(* IEC 61131-3 sources: daoli-st-library/DL_MathData (part 25) *)

(* ---- FC_DL_StringReplaceAtEx.st ---- *)
(*
    FC_DL_StringReplaceAtEx —— 定位定长替换防御包装（与 StringReplaceAll 全局替换职责区分）
    ------------------------------------------------------------------
    分类      : DL_MathData / String
    前缀      : FC_DL_
    版本      : 1.0.0
    溯源      : IEC 61131-3 标准语义的道莅防御性实现
                （内部委托平台内建函数，外围统一错误码/钳位/双语文档；
                  未复制任何闭源厂商源码，参考实现仅限 MIT/Apache 许可）
    平台      : 纯 IEC 61131-3，CODESYS / TwinCAT / InoProShop 通用
    作者      : 道莅代码库 · PLC编程专家（R15）
    ------------------------------------------------------------------
    功能说明  : 与既有 FC_DL_StringReplaceAll（全串搜索全局替换）职责明
                确区分：本件为定位置定长覆盖——自 nPos 位序（1 基）起用
                sRep 覆盖，不搜索、不改变总长，sRep 超出串尾部分被截断。
                nPos < 1 钳 1 置 16#0001_01BD；nPos > len 原样返回置 16#0001_01BD；覆盖长
                度 = MIN(sRep 长, len-nPos+1)，sRep 被截断时按 R37 范式显
                式置 bTruncated=TRUE 与 16#0001_028B。先整串复制再覆盖（各轮带
                255 越界 EXIT 守卫），复制后显式写空字符终止符。返回值
                TRUE 表示已执行完成。
    错误码    : 0000 正常 / 16#0001_01BD 入参越界（nPos 钳位或超串长，超长时原样返回） / 16#0001_028B 上溢下溢（sRep 超串尾被截断，bTruncated=TRUE）
    修订记录  : 2026-11-16 v1.0.0 首次入库（R15）
*)
FUNCTION FC_DL_StringReplaceAtEx : BOOL
VAR_INPUT
    sIn  : STRING(255); // 源串 [字符] / source string [chars]
    sRep : STRING(255); // 覆盖串 [字符]，超串尾部分被截断 / replacement string [chars], tail beyond the source end truncated
    nPos : INT; // 覆盖起始位序 [字符位序]，1 基 / overwrite start position [char position], 1-based
END_VAR
VAR_OUTPUT
    sResult    : STRING(255); // 结果串 [字符]，总长与源串一致 / result string [chars], same length as the source
    eErr : UDINT; // 错误码，0=正常，1=位置钳位/超长，2=覆盖串截断 / error id, 0=ok, 1=position clamped or beyond length, 2=replacement truncated
    bError     : BOOL; // 是否出错，eErr 非 0 时为 TRUE / error flag, TRUE when eErr is nonzero
    bValid     : BOOL; // 输出是否有效可用 / output valid
    bTruncated : BOOL; // 截断标志，sRep 超串尾被截断时 TRUE（R37 范式） / truncation flag, TRUE when the replacement was tail-truncated
END_VAR
VAR
    nI      : INT; // 循环索引 [字符位序]，1 基 / loop index [char position], 1-based
    nLen    : INT; // 锁存的源串有效长度 [字符] / latched effective source length [chars]
    nRepLen : INT; // 锁存的覆盖串有效长度 [字符] / latched effective replacement length [chars]
    nPosC   : INT; // 钳位后的覆盖起始位序 [字符位序] / clamped overwrite start position [char position]
    nAvail  : INT; // 自起点起可用字符数 [字符] / chars available from the start position [chars]
    nUseRep : INT; // 覆盖串实际复制数 [字符] / chars actually copied from the replacement [chars]
END_VAR
VAR CONSTANT
    DL_RA_MAX : INT := 255; // 串型上限 [字符] / string type cap [chars]
END_VAR

// 段 1｜返回值与输出预置，任何早退路径不留脏码 / segment 1, preset return value and outputs
FC_DL_StringReplaceAtEx := TRUE; // 返回值预置 TRUE（已执行口径） / preset return to TRUE
sResult                 := ''; // 结果串预置空串 / preset result to the empty string
eErr                := 16#0000_0000; // 错误码预置正常 / preset error id to ok
bError                  := FALSE; // 错误标志预置无错 / preset error flag to FALSE
bValid                  := TRUE; // 有效标志预置可用 / preset valid flag to TRUE
bTruncated              := FALSE; // 截断标志预置无截断 / preset truncation flag to FALSE

// 段 2｜两串有效长度各一次锁存（空字符截止扫描 + 255 越界守卫） / segment 2, latch both effective lengths once
nI      := 1; // 索引起始 [字符位序] / index start
nLen    := 0; // 源串长度预置 [字符] / preset source length
WHILE nI <= DL_RA_MAX DO
    IF nI > DL_RA_MAX THEN    (* 越界守卫（双重保险） EN: overrun guard *)
        EXIT;
    END_IF
    IF sIn[nI] = '$00' THEN   (* 首个空字符即串结束 EN: first null char ends the string *)
        EXIT;
    END_IF
    nLen := nI; // 记录源串最后非空位序 [字符] / record the last non-null position
    nI   := nI + 1; // 每轮自增 / per-iteration increment
END_WHILE
nI      := 1; // 索引复位 / reset index
nRepLen := 0; // 覆盖串长度预置 [字符] / preset replacement length
WHILE nI <= DL_RA_MAX DO
    IF nI > DL_RA_MAX THEN    (* 越界守卫（双重保险） EN: overrun guard *)
        EXIT;
    END_IF
    IF sRep[nI] = '$00' THEN  (* 首个空字符即串结束 EN: first null char ends the string *)
        EXIT;
    END_IF
    nRepLen := nI; // 记录覆盖串最后非空位序 [字符] / record the last non-null position
    nI      := nI + 1; // 每轮自增 / per-iteration increment
END_WHILE

// 段 3｜位置闸门：nPos < 1 钳 1 置 16#0001_01BD；nPos > len 原样返回置 16#0001_01BD / segment 3, position gate, below 1 clamped to 1, beyond length returns the original with code 1
IF nPos < 1 THEN
    nPosC := 1; // 下越界钳 1 / clamped to 1
    eErr := 16#0001_01BD; // 入参越界码 / out-of-domain code
    bError   := TRUE; // 置错误标志 / raise error flag
    bValid   := FALSE; // 钳位降级 / degraded output
ELSE
    nPosC := nPos; // 域内直通 / in-domain pass-through
END_IF
IF nPosC > nLen THEN
    FOR nI := 1 TO nLen DO
        IF nI > DL_RA_MAX THEN   (* 越界守卫（双重保险） EN: overrun guard *)
            EXIT;
        END_IF
        sResult[nI] := sIn[nI]; // 位置超长原样返回 / position beyond length, original returned
    END_FOR
    IF nLen < DL_RA_MAX THEN
        sResult[nLen + 1] := '$00'; // 空字符终止符 / null terminator
    END_IF
    eErr := 16#0001_01BD; // 入参越界码（首事件优先不覆盖钳位码） / out-of-domain code, first event kept
    bError   := TRUE; // 置错误标志 / raise error flag
    bValid   := FALSE; // 输出不可用 / output invalid
    RETURN;
END_IF

// 段 4｜覆盖配额闸（R37 范式：先判定后写入，严禁静默回夹） / segment 4, overwrite quota gate, R37 paradigm, decide before writing
nAvail := nLen - nPosC + 1; // 自起点起可用字符数 [字符] / chars available from the start
IF nRepLen > nAvail THEN
    nUseRep := nAvail; // 覆盖串截到串尾 / replacement clipped to the string end
    bTruncated := TRUE; // 显式置截断标志（R37 教训） / set the truncation flag explicitly
    eErr   := 16#0001_028B; // 上溢码：sRep 超串尾已截断 / overflow code, replacement tail-truncated
    bError     := TRUE; // 置错误标志 / raise error flag
    bValid     := FALSE; // 截断降级结果 / degraded truncated output
ELSE
    nUseRep := nRepLen; // 域内直通 / in-domain pass-through
END_IF

// 段 5｜整串复制：FOR 循环 + 255 越界 EXIT 守卫 / segment 5, copy the whole source with the overrun guard
FOR nI := 1 TO nLen DO
    IF nI > DL_RA_MAX THEN       (* 越界守卫（双重保险） EN: overrun guard *)
        EXIT;
    END_IF
    sResult[nI] := sIn[nI]; // 逐字符复制 / char-by-char copy
END_FOR

// 段 6｜定长覆盖：目的位序 = nPos 起顺延，超 255 即退出 / segment 6, fixed-position overwrite
FOR nI := 1 TO nUseRep DO
    IF (nPosC + nI - 1) > DL_RA_MAX THEN   (* 目的侧越界守卫 EN: destination overrun guard *)
        EXIT;
    END_IF
    IF nI > DL_RA_MAX THEN                 (* 源侧越界守卫 EN: source overrun guard *)
        EXIT;
    END_IF
    sResult[nPosC + nI - 1] := sRep[nI]; // 逐字符覆盖 / char-by-char overwrite
END_FOR

// 段 7｜显式写终止符：总长与源串一致 / segment 7, write the terminator explicitly, total length equals the source
IF nLen < DL_RA_MAX THEN
    sResult[nLen + 1] := '$00'; // 空字符终止符 / null terminator
END_IF
END_FUNCTION

(* ---- FC_DL_StringRightEx.st ---- *)
(*
    FC_DL_StringRightEx —— 取右 n 字符防御包装（n 越界钳位 + 255 守卫逐字符复制）
    ------------------------------------------------------------------
    分类      : DL_MathData / String
    前缀      : FC_DL_
    版本      : 1.0.0
    溯源      : IEC 61131-3 标准语义的道莅防御性实现
                （内部委托平台内建函数，外围统一错误码/钳位/双语文档；
                  未复制任何闭源厂商源码，参考实现仅限 MIT/Apache 许可）
    平台      : 纯 IEC 61131-3，CODESYS / TwinCAT / InoProShop 通用
    作者      : 道莅代码库 · PLC编程专家（R15）
    ------------------------------------------------------------------
    功能说明  : 取源串右侧 nCount 个字符到 sResult。采用逐字符 FOR 复制
                （跨平台口径，不依赖平台 RIGHT 行为差异），源/目的双侧
                均带 255 越界 EXIT 守卫，复制后显式写空字符终止符。
                nCount <= 0 返回空串置 16#0001_01A6；nCount > 实际长度返回全串并
                置 16#0001_01A4（bValid=FALSE，截断诉求由错误码显式体现）。返回值
                TRUE 表示函数已执行完成，结果总在 sResult 中。
    错误码    : 0000 正常 / 16#0001_01A4 入参越界（nCount 超实际长度，已返回全串） / 16#0001_01A6 无效入参（nCount <= 0）
    修订记录  : 2026-11-16 v1.0.0 首次入库（R15）
*)
FUNCTION FC_DL_StringRightEx : BOOL
VAR_INPUT
    sIn    : STRING(255); // 源串 [字符] / source string [chars]
    nCount : INT; // 请求取右字符数 [字符]，<= 0 判无效 / requested right char count [chars], values at or below 0 invalid
END_VAR
VAR_OUTPUT
    sResult  : STRING(255); // 结果串 [字符]，右 nCount 字符 / result string [chars], right nCount chars
    eErr : UDINT; // 错误码，0=正常 / error id, 0=ok
    bError   : BOOL; // 是否出错，eErr 非 0 时为 TRUE / error flag, TRUE when eErr is nonzero
    bValid   : BOOL; // 输出是否有效可用 / output valid
END_VAR
VAR
    nI      : INT; // 循环索引 [字符位序]，1 基 / loop index [char position], 1-based
    nLen    : INT; // 锁存的源串有效长度 [字符] / latched effective source length [chars]
    nUse    : INT; // 实际复制字符数 [字符] / chars actually copied [chars]
    nSrcBgn : INT; // 源串复制起点 [字符位序] / source copy start position [char position]
END_VAR
VAR CONSTANT
    DL_RT_MAX : INT := 255; // 串型上限 [字符] / string type cap [chars]
END_VAR

// 段 1｜返回值与输出预置，任何早退路径不留脏码 / segment 1, preset return value and outputs
FC_DL_StringRightEx := TRUE; // 返回值预置 TRUE（已执行口径） / preset return to TRUE, executed semantics
sResult             := ''; // 结果串预置空串 / preset result to the empty string
eErr            := 16#0000_0000; // 错误码预置正常 / preset error id to ok
bError              := FALSE; // 错误标志预置无错 / preset error flag to FALSE
bValid              := TRUE; // 有效标志预置可用 / preset valid flag to TRUE

// 段 2｜源串有效长度一次锁存（空字符截止扫描 + 255 越界守卫） / segment 2, latch the effective source length once
nI   := 1; // 索引起始 [字符位序] / index start
nLen := 0; // 有效长度预置 [字符] / preset effective length
WHILE nI <= DL_RT_MAX DO
    IF nI > DL_RT_MAX THEN   (* 越界守卫（双重保险） EN: overrun guard, defense in depth *)
        EXIT;
    END_IF
    IF sIn[nI] = '$00' THEN  (* 首个空字符即串结束 EN: first null character marks the string end *)
        EXIT;
    END_IF
    nLen := nI; // 记录最后非空字符位序 [字符] / record the last non-null char position
    nI   := nI + 1; // 每轮自增 / per-iteration increment
END_WHILE

// 段 3｜入参域闸门：nCount <= 0 无效置 16#0001_01A6；nCount 超长度钳到全长置 16#0001_01A4 / segment 3, input domain gate
IF nCount <= 0 THEN
    sResult  := ''; // 无效入参返回空串 / invalid input returns the empty string
    eErr := 16#0001_01A6; // 无效入参码 / invalid input code
    bError   := TRUE; // 置错误标志 / raise error flag
    bValid   := FALSE; // 输出不可用 / output invalid
    RETURN;
ELSIF nCount > nLen THEN
    nUse    := nLen; // 请求超长，钳到全串长 / request beyond length, clamped to full length
    eErr := 16#0001_01A4; // 入参越界码：截断诉求显式置码 / out-of-domain code, truncation intent made explicit
    bError   := TRUE; // 置错误标志 / raise error flag
    bValid   := FALSE; // 输出为截断降级结果 / output is a degraded truncated result
ELSE
    nUse := nCount; // 域内直通 / in-domain pass-through
END_IF
nSrcBgn := nLen - nUse + 1; // 源串复制起点 = 长度减取数加一 [字符位序] / source start = length minus count plus one

// 段 4｜逐字符复制（跨平台口径）：源/目的双侧 255 越界 EXIT 守卫 / segment 4, char-by-char copy with overrun guards on both source and destination
FOR nI := 1 TO nUse DO
    IF nI > DL_RT_MAX THEN            (* 目的侧越界守卫 EN: destination overrun guard *)
        EXIT;
    END_IF
    IF (nSrcBgn + nI - 1) > DL_RT_MAX THEN   (* 源侧越界守卫 EN: source overrun guard *)
        EXIT;
    END_IF
    sResult[nI] := sIn[nSrcBgn + nI - 1]; // 逐字符复制 / char-by-char copy
END_FOR

// 段 5｜显式写终止符 / segment 5, write the terminator explicitly
IF nUse < DL_RT_MAX THEN
    sResult[nUse + 1] := '$00'; // 空字符终止符 / null terminator
END_IF
END_FUNCTION

(* ---- FC_DL_StringSplit.st ---- *)
(*==============================================================================
 * 组件名称 (Component)  : FC_DL_StringSplit
 * 所属子库 (Sublibrary) : DL_MathData
 * 当前版本 (Version)    : 1.0.0
 * 兼容性   (Platform)   : CODESYS 3.5 / TwinCAT 3 / 汇川 InoProShop / Machine Expert
 *                         仅依赖 Standard.library 的标准串函数（LEN / FIND / LEFT / DELETE）
 * 功能描述 (Function)   : 按单字符分隔符把报文拆分为字段数组。返回实际拆分出的字段数，
 *                         字段写入调用方提供的持久数组（引用型输入输出）。
 *                         采用"定位 → 取字段 → 吃掉已处理段"的标准循环，全库统一口径，
 *                         替代各项目各写一套的重复劳动（主流平台均无内置拆分函数）。
 *                         相邻分隔符产生空字段，符合 CSV 语义，不跳过、不合并；
 *                         字段数超出调用方上限时，剩余整段并入末字段并置截断标志，
 *                         结果不静默丢弃。
 * 开源溯源 (Origin)     : 原创实现。定位取段的处理范式为公开通行做法；
 *                         空字段语义与截断语义为本库差异化设计，未复制任何源码。
 * 本文件内含       : FC    FC_DL_StringSplit（单 POU，无配套类型）
 * 依赖     (Depends)    : 无 DL_ 内部依赖；Standard.library: LEN / FIND / LEFT / DELETE
 * 红线自检 (Redline)    : R1 ✓ 禁用全局存储与物理寻址 ｜ R2 ✓ 无地址直写
 *                         R3 ✓ 仅标准串函数 ｜ R4 ✓ 主循环防死锁 + 字段数钳位 + 下标双检
 *                         R5 ✓ 全变量中英双语同行注释 ｜ R6 N/A（纯函数，无状态机）
 *                         R7 N/A（无定时器/边沿实例）｜ R8 ✓ 字段上限与循环上限全常量化
 *
 * 【输出缓冲纪律 / Output buffer discipline（边界 B7，反例警告）】
 *   字段数组为引用型输入输出，调用方必须传入持久数组并在每次调用前自行清场。
 *   反例：把临时变量或每次新构造的数组传进来，上一次调用的残留字段会留在数组里，
 *   本次字段数变少时旧字段仍然可见，表现为"配方里凭空多出几个字段"的诡异故障。
 *   正确做法：一个报文一个专用数组，调用前用循环把数组元素清成空串。
 *
 * 【内存要求 / Memory requirement（边界 B10）】
 *   调用方需持有 16 × 256 字节约 4KB 的字段缓冲。单次调用最坏 16 次定位/取段/删除，
 *   无嵌套循环，耗时与报文长度呈线性关系。
 *
 * 【单字符锁定 / Single-character delimiter（边界 B1，决策 D-R2-18）】
 *   分隔符长度必须恰好为 1，否则直接拒绝且不拆分。多字符分隔会同时复杂化
 *   定位语义与截断语义，单字符已覆盖 CSV / 分号 / 竖线全部主流场景。
 *
 * 修订历史 (Revision)   :
 *   2026-11-14  v1.0.0  首版入库（Phase 1 第二轮 · Level 0 批次 A）
 *============================================================================*)
FUNCTION FC_DL_StringSplit : INT
VAR_INPUT
    sSource    : STRING(255);                 // 待拆分报文，最大 255 字符 / Source message, 255 characters max
    sDelimiter : STRING(1) := ',';            // 分隔符（单字符） / Single-character delimiter
    uMaxFields : INT := 16;                   // 最大输出字段数 [个]，合法域 1..16 / Max output fields [count], valid 1..16
END_VAR
VAR_IN_OUT
    aFields    : ARRAY[0..15] OF STRING(255); // 输出字段缓冲，调用方持有并复用 / Caller-owned reusable output buffer
END_VAR
VAR_OUTPUT
    bValid     : BOOL;                        // 拆分完整标志，FALSE = 发生截断 / Complete flag, FALSE = truncated
    uErrorId   : UDINT;                       // 故障码，0 = 无故障 / Error code, 0 = no error
END_VAR
VAR
    sTmp       : STRING(255);   // 剩余段工作副本，源串全程只读 / Working copy of the remaining segment
    nDelimPos  : INT;           // 分隔符位置（1 起始，0 = 未找到） / Delimiter position, 1-based, 0 = not found
    nFieldIdx  : INT;           // 当前字段索引 [个] / Current field index [count]
    nFieldLen  : INT;           // 当前字段长度 [字符] / Current field length [characters]
    nDelimLen  : INT;           // 分隔符长度校验值 [字符] / Delimiter length check value [characters]
    nMaxEff    : INT;           // 钳位后的最大字段数 [个] / Clamped max fields [count]
    nSrcLen    : INT;           // 源串有效长度 [字符] / Effective source length [characters]
    bRun       : BOOL;          // 循环继续标志 / Loop continuation flag
    nGuard     : DINT;          // 循环防死锁计数器 [次] / Loop deadlock guard counter [count]
    nLoop      : INT;           // 主循环索引 [次] / Main loop index [count]
END_VAR
VAR CONSTANT
    DL_SP_MAX_FIELDS : INT  := 16;   // 字段数上限 [个]，与数组维度一致 / Field cap [count], must match the array
    DL_SP_LOOP_MAX   : DINT := 64;   // 主循环防死锁上限 [次]，字段数 × 余量 / Loop guard limit [count]
    DL_SP_LEN_MAX    : INT  := 255;  // 报文字符上限 [字符]，与类型声明一致 / Message length cap [characters]
END_VAR

(*------------------------------------------------------------------------------
 * 段 1｜结果预置（P-01 范式）：先给 0 字段与成功标志
 *      Safe preset: zero fields and a success flag
 *-----------------------------------------------------------------------------*)
FC_DL_StringSplit := 0;
bValid   := TRUE;
uErrorId := 16#0000_0000;
nFieldIdx := 0;
nFieldLen := 0;
nMaxEff   := uMaxFields;

(*------------------------------------------------------------------------------
 * 段 2｜分隔符合法性（边界 B1）：长度不为 1 直接拒绝，不进入拆分流程
 *      Delimiter validity: any length other than one is rejected before splitting
 *-----------------------------------------------------------------------------*)
nDelimLen := LEN(sDelimiter);

IF nDelimLen <> 1 THEN
    bValid   := FALSE;
    uErrorId := 16#0001_0008;
    FC_DL_StringSplit := 0;
ELSE

    (*--------------------------------------------------------------------------
     * 段 3｜字段数钳位（边界 B2）：越界钳位后继续拆分，不停机
     *      Field count clamping: clamp and keep splitting, never stop the machine
     *-------------------------------------------------------------------------*)
    IF nMaxEff < 1 THEN
        nMaxEff  := 1;
        uErrorId := 16#0001_0001;
    ELSIF nMaxEff > DL_SP_MAX_FIELDS THEN
        nMaxEff  := DL_SP_MAX_FIELDS;
        uErrorId := 16#0001_0001;
    END_IF

    (* 源串长度先钳位再用：超长报文的尾部按截断处理，绝不越界读 *)
    (* Source length clamped first: an over-length message is treated as truncated *)
    nSrcLen := LEN(sSource);
    IF nSrcLen > DL_SP_LEN_MAX THEN
        nSrcLen := DL_SP_LEN_MAX;
    ELSIF nSrcLen < 0 THEN
        nSrcLen := 0;
    END_IF

    IF nSrcLen = 0 THEN
        (* 空源串是合法结果而非错误（边界 B3） *)
        (* An empty source is a legal result, not an error *)
        FC_DL_StringSplit := 0;
    ELSE

        (*----------------------------------------------------------------------
         * 段 4｜主循环（边界 B4/B5/B6）：定位、取段、删除已处理段
         *      Main loop: locate, extract, then drop the handled prefix
         *      已到最后一个可用字段而串内仍有分隔符时，剩余整段并入末字段并置截断标志
         *      On the last usable field with delimiters left, the whole remainder is kept
         *      并在置位截断标志，调用方据此识别"字段没拆完"
         *      and the truncation flag is raised so the caller can tell fields were cut
         *---------------------------------------------------------------------*)
        sTmp   := sSource;
        nLoop  := 0;
        bRun   := TRUE;
        nGuard := 0;

        WHILE bRun DO

            IF nFieldIdx >= nMaxEff THEN
                bRun := FALSE;
            ELSE
                nDelimPos := FIND(sTmp, sDelimiter);

                IF (nDelimPos > 0) AND ((nFieldIdx + 1) < nMaxEff) THEN
                    (*----------------------------------------------------------
                     * 段 4a｜常规切分：字段 = 分隔符之前的部分，然后吃掉分隔符
                     *      Normal split: the field precedes the delimiter, which is dropped
                     *      连续分隔符会自然产生长度为 0 的空字段，不跳过（边界 B6）
                     *      Consecutive delimiters yield empty fields, never skipped
                     *---------------------------------------------------------*)
                    nFieldLen := nDelimPos - 1;

                    IF nFieldLen < 0 THEN
                        nFieldLen := 0;
                    END_IF

                    IF (nFieldIdx >= 0) AND (nFieldIdx < DL_SP_MAX_FIELDS) THEN
                        aFields[nFieldIdx] := LEFT(sTmp, nFieldLen);
                    END_IF

                    sTmp      := DELETE(sTmp, nDelimPos, nDelimLen);
                    nFieldIdx := nFieldIdx + 1;

                ELSE
                    (*----------------------------------------------------------
                     * 段 4b｜末段落地：无分隔符，或已到最后一个可用字段
                     *      Final segment: no delimiter left, or the last usable field
                     *      后者若串内仍有分隔符即为截断，剩余整段并入末字段并告警
                     *      The latter with a delimiter present is a truncation and is flagged
                     *---------------------------------------------------------*)
                    IF (nFieldIdx >= 0) AND (nFieldIdx < DL_SP_MAX_FIELDS) THEN
                        aFields[nFieldIdx] := sTmp;
                    END_IF

                    nFieldIdx := nFieldIdx + 1;

                    IF nDelimPos > 0 THEN
                        bValid   := FALSE;
                        uErrorId := 16#0001_000D;
                    END_IF

                    sTmp := '';
                    bRun := FALSE;
                END_IF

            END_IF

            (* 防死锁：每轮字段索引必然递增，仍设上限兜底防止异常串函数导致死循环 *)
            (* Deadlock guard: the index always advances, the cap is a second line of defence *)
            nGuard := nGuard + 1;
            nLoop  := nLoop + 1;

            IF (nGuard > DL_SP_LOOP_MAX) OR (nLoop > DL_SP_MAX_FIELDS) THEN
                bRun     := FALSE;
                bValid   := FALSE;
                IF uErrorId = 16#0000_0000 THEN
                    uErrorId := 16#0001_0004;
                END_IF
            END_IF

        END_WHILE;

        (*----------------------------------------------------------------------
         * 段 5｜返回值：实际字段数，异常路径返回已完成的数量（P-01）
         *      Return value: the actual field count, partial counts on abnormal paths
         *---------------------------------------------------------------------*)
        IF nFieldIdx < 0 THEN
            FC_DL_StringSplit := 0;
        ELSIF nFieldIdx > DL_SP_MAX_FIELDS THEN
            FC_DL_StringSplit := DL_SP_MAX_FIELDS;
        ELSE
            FC_DL_StringSplit := nFieldIdx;
        END_IF

    END_IF
END_IF
END_FUNCTION

(* ---- FC_DL_StringStripCharsEx.st ---- *)
(*==============================================================================
 * 组件名称 (Component)  : FC_DL_StringStripCharsEx
 * 所属子库 (Sublibrary) : DL_MathData
 * 归属目录 (Directory)  : C:\Library\DL_MathData
 * 当前版本 (Version)    : 1.0.0
 * 分类/来源标签         : 函数（FUNCTION）· 纯函数 · 自定义字符集剥离
 *                         iec-std-wrapper / string / r37-reference
 * 兼容性   (Platform)   : CODESYS 3.5 / TwinCAT 3 / 汇川 InoProShop / 施耐德
 *                         Machine Expert；仅用 Standard.library 的 LEN / MID / FIND
 * 溯源声明 (Provenance) : IEC 61131-3 标准语义的道莅防御性实现——内部委托平台标准库语义，
 *                         外围统一错误码 / 钳位 / 双语注释，严禁重实现数学内核。
 * 功能一句话 (Summary)  : 去除字符串两侧属于自定义字符集的字符（区别于仅去空格的
 *                         Trim），空集输入恒等返回，全程 R37 四步长度守卫。
 *
 * 功能描述 (Function)   : LEN 一次锁存源长并与 255 比较，超限按 bAllowTrunc 分路；
 *                         合法路径用 FIND 判字符归属，从左向右收缩首界、从右向左
 *                         收缩尾界，中段一次 MID 取出，出口做长度一致性校验。
 * 与既有件边界 (Boundary): FC_DL_StringTrim 只去空格且语义固定；本件字符集是契约
 *                         参数，空串字符集即为恒等变换，不做任何猜测性补剥离。
 * 码位说明 (Codes)      : 信息 16#0002_3038 有剥离发生（nStripped 大于零）
 *                         故障 16#0002_3039 源长度域外且未允许截断（防御闸）
 *                         故障 16#0002_303A 中段取出长度与预期不一致（防御校验）
 *                         段 16#02_3_38~3B 首槽信息级、次槽起故障级。
 * 依赖说明 (Depends)    : 无 DL_ 内部依赖；仅 Standard.library 的 LEN / MID / FIND。
 * 镜像量清单 (R38)      : nSrcLen 唯一锁存量；nFirst 与 nLast 是本件的两个消费边界，
 *                         中段长度 nKeep 全部由该副本与两界导出，不重复取 LEN。
 * 红线自检 (Redline)    : 零全局依赖 ｜ 零 VAR_EXTERNAL ｜ 零 %I/%Q ｜ 纯 IEC 标准库
 *                         无除法故无除零面 ｜ 全变量双语同行注释 ｜ 无定时器实例
 * 修订历史 (Revision)   : 2026-11-18  v1.0.0  首版入库（R32 · 批 1）
 *============================================================================*)

FUNCTION FC_DL_StringStripCharsEx : BOOL
VAR_INPUT
    sSrc        : STRING(255);      // 源文本 [ASCII]，定长 255 / Source text, fixed 255 characters
    sStrip      : STRING(255);      // 剥离字符集 [ASCII]，空串即恒等 / Strip charset, empty means identity
    bAllowTrunc : BOOL := FALSE;    // 允许截断，真则截断写出，假则拒绝构造 / TRUE truncates and writes, FALSE refuses
END_VAR
VAR_OUTPUT
    sOut        : STRING(255);      // 剥离结果 [ASCII] / Stripped result
    bTruncated  : BOOL;             // 截断标志，源超上限时为真 / Set true when the source exceeded the limit
    nStripped   : INT;              // 两侧剥离的字符总数 [个] / Total characters stripped from both ends
    uErrorId    : UDINT;            // 事件码，0 表示无事件 / Event code, zero means none
END_VAR
VAR
    sMid     : STRING(255); // 中段暂存 [ASCII] / Middle segment staging
    cCh      : STRING(1);   // 当前字符 [字符] / Current character
    nSrcLen  : INT;         // 锁存的源文本长度 [字符]，R38 唯一锁存量 / Latched source length
    nFirst   : INT;         // 左边界，1 起 [索引] / Left boundary, 1-based
    nLast    : INT;         // 右边界 [索引] / Right boundary
    nKeep    : INT;         // 中段长度 [字符] / Middle segment length
    uCode    : UDINT;       // 码位暂存，出口单点写入 [码] / Code staging
END_VAR
VAR CONSTANT
    DL_STS_MAXLEN : INT := 255; // 字符串上限 [字符]，与形参声明一致 / String limit, matches the declarations
    DL_STS_ONE    : INT := 1;   // 单字符长度参数 [字符] / Single character length argument
END_VAR

(* 段 1｜输出预置与残留清除 / Pre-set and clear before any branch *)
FC_DL_StringStripCharsEx := FALSE;
sOut       := '';
sMid       := '';
bTruncated := FALSE;
nStripped  := 0;
uErrorId   := 16#0000_0000;
uCode      := 16#0000_0000;

(* 段 2｜R37 第 1 步：LEN 一次锁存 / Step one: latch the length once *)
nSrcLen := LEN(sSrc);
IF nSrcLen < 0 THEN
    nSrcLen := 0;                // 防御：异常返回值钳到零 / Defensive: clamp an anomalous result
END_IF

(* 段 3｜R37 第 2、3 步：与上限比较，超限先置标志后分路 / Compare, flag first, then branch *)
IF nSrcLen > DL_STS_MAXLEN THEN
    bTruncated := TRUE;          // 事实先记录 / Record the fact first
    IF NOT bAllowTrunc THEN
        uErrorId := 16#0002_3039; // 故障级：拒绝构造 / Fault: refuse to build
        RETURN;
    END_IF
    nSrcLen := DL_STS_MAXLEN;    // 第 4 步截断路 / Truncation path
END_IF

(* 段 4｜左界收缩：首字符属于字符集则右移 / Shrink the left boundary while the first char belongs to the set *)
nFirst := 1;
WHILE (nFirst <= nSrcLen) DO
    cCh := MID(sSrc, DL_STS_ONE, nFirst);            // 取当前首字符 / Take the current first character
    IF FIND(sStrip, cCh) > 0 THEN
        nFirst := nFirst + DL_STS_ONE;               // 属集，右移 / Belongs, shift right
    ELSE
        EXIT;                                        // 非属，停 / Not belonging, stop
    END_IF
END_WHILE

(* 段 5｜右界收缩：尾字符属于字符集则左移，越左界即停 / Shrink the right boundary, stop at the left one *)
nLast := nSrcLen;
WHILE (nLast >= nFirst) DO
    cCh := MID(sSrc, DL_STS_ONE, nLast);             // 取当前尾字符 / Take the current last character
    IF FIND(sStrip, cCh) > 0 THEN
        nLast := nLast - DL_STS_ONE;                 // 属集，左移 / Belongs, shift left
    ELSE
        EXIT;                                        // 非属，停 / Not belonging, stop
    END_IF
END_WHILE

(* 段 6｜中段一次取出：长度由两界导出，空段显式置空串 / Take the middle once; an empty segment is explicitly empty *)
nKeep := nLast - nFirst + DL_STS_ONE;                // 中段长度导出 / Derive the middle length
IF nKeep < 0 THEN
    nKeep := 0;                  // 结构性非负，仍显式兜底 / Structurally non-negative, belt and braces
END_IF
IF nKeep > 0 THEN
    sMid := MID(sSrc, nKeep, nFirst);                // 一次取出中段 / Take the middle in one shot
ELSE
    sMid := '';                  // 全串被剥离，结果空串 / Whole string stripped, result empty
END_IF

(* 段 7｜写出一致性校验（防御闸）与出口装配 / Write consistency gate and exit assembly *)
IF LEN(sMid) <> nKeep THEN
    uErrorId := 16#0002_303A;    // 故障级：取出链路异常，结果作废 / Fault: extraction chain broken
    sOut := '';
    RETURN;
END_IF
nStripped := nSrcLen - nKeep;    // 剥离计数导出 / Derive the stripped count
IF nStripped > 0 THEN
    uCode := 16#0002_3038;       // 信息级：有剥离发生 / Info: stripping happened
END_IF
sOut := sMid;
uErrorId := uCode;               // 码位单点写入 / Single write point for the code
FC_DL_StringStripCharsEx := TRUE;
END_FUNCTION

(* ---- FC_DL_StringToLowerEx.st ---- *)
(*==============================================================================
 * 组件名称 (Component)  : FC_DL_StringToLowerEx
 * 所属子库 (Sublibrary) : DL_MathData
 * 归属目录 (Directory)  : C:\Library\DL_MathData
 * 当前版本 (Version)    : 1.0.0
 * 分类/来源标签         : 函数（FUNCTION）· 纯函数 · 字符串小写扩展转换
 *                         iec-std-wrapper / string / r40-reference
 * 兼容性   (Platform)   : CODESYS 3.5 / TwinCAT 3 / 汇川 InoProShop / 施耐德
 *                         Machine Expert；仅用 Standard.library 的 LEN / MID / CONCAT / FIND
 * 溯源声明 (Provenance) : IEC 61131-3 标准语义的道莅防御性实现——内部委托平台标准库语义，
 *                         外围统一错误码 / 钳位 / 双语注释，严禁重实现数学内核。
 * 功能一句话 (Summary)  : 把 ASCII 域内大写字母映射为小写，域外字符保持原值并计数，
 *                         超长按截断标志显式分路，空串原样直通。
 * 本件存在的意义 (Why this unit exists)：
 *   各平台自带的大小写转换行为不一（有的吞掉高位字符、有的整串拒绝），本件只用
 *   标准 LEN/MID/CONCAT/FIND 做逐字符查表映射：大写字母经双码表定位转小写，
 *   其余字符原样保留并以信息码告知「有保留发生」，调用方永远知道结果里混了什么。
 * 功能描述 (Function)   : 第 1 步 LEN 一次锁存源长；第 2 步与 255 上限比较；第 3 步
 *                         超限先置截断标志（255 上限显式化，不依赖平台隐式截断）；
 *                         第 4 步按 bAllowTrunc 分路截断写出或拒绝。
 *                         空串直通：源长为 0 时不进循环、写出计数 0 等于源长 0，
 *                         出口装配返回 TRUE 且不占任何码位。
 *                         合法路径逐字符取字符：落在 'A'..'Z' 域内的用 FIND 在大写
 *                         码表定位后到同位小写码表取字符，域外字符保持并累计 nKept。
 * 与既有件边界 (Boundary): 本件为 FC_DL_StringToUpperEx 的严格对偶件（映射方向互逆、
 *                         四步样板与分路口径逐条对应），只做 ASCII A..Z 域内映射，
 *                         不做 Unicode 与本地化。
 * 码位说明 (Codes)      : 信息 16#0001_0499 源超 255 上限，已按上限截断写出
 *                         故障 16#0001_03D4 源超上限且未允许截断（防御闸拒绝）
 *                         故障 16#0001_03D5 写出计数与源长不一致（防御校验）
 *                         （R90 反证句：截断事实无法由 sDst 观测——截断与正常写出
 *                           结果均为合法串且返回值同为 TRUE，故截断侧须占码；
 *                           计数不一致属写出链路异常，与截断、保留场景的输出组合
 *                           （空串加故障码）均不同，故独立占码）
 * 依赖说明 (Depends)    : 无 DL_ 内部依赖；仅 Standard.library 的 LEN / MID / CONCAT / FIND。
 * 镜像量清单 (R38)      : nSrcLen 是本件唯一锁存量，入口一次导出，其后比较与循环
 *                         上界全部读该副本，全文不再对入参串取长度。
 * 遗留假设 (Legacy)     : 字符比较使用 >= / <= 排序比较（与库内 FC_DL_StringToUpperEx
 *                         同口径）；若某平台未实现 STRING 排序比较，须在编译门槛里
 *                         核对后改走 FIND 查表判定。
 * 红线自检 (Redline)    : 零全局依赖 ｜ 零 VAR_EXTERNAL ｜ 零 %I/%Q ｜ 纯 IEC 标准库
 *                         无除法故无除零面 ｜ 全变量双语同行注释 ｜ 无定时器实例
 * 修订历史 (Revision)   : 2026-11-19  v1.0.0  首版入库（R40 · 批 3 · T0 快车道）
 *============================================================================*)

FUNCTION FC_DL_StringToLowerEx : BOOL
VAR_INPUT
    sSrc        : STRING(255);      // 源文本 [ASCII]，定长 255 ｜ source text, fixed 255 characters
    bAllowTrunc : BOOL := FALSE;    // 允许截断，真则截断写出，假则拒绝构造 ｜ TRUE truncates and writes, FALSE refuses
END_VAR
VAR_OUTPUT
    sDst        : STRING(255);      // 小写结果 [ASCII]，域外字符保持原值 ｜ lowercase result, out-of-domain chars kept
    bTruncated  : BOOL;             // 截断标志，源超上限时为真 ｜ set true when the source exceeded the limit
    nKept       : INT;              // 保持原值的域外字符个数 [个] ｜ count of kept out-of-domain characters
    uErrorId    : UDINT;            // 事件码，0 表示无事件 ｜ event code, zero means none
END_VAR
VAR
    sTmp     : STRING(255); // 结果累积缓冲 [ASCII]，出口一次性赋给 sDst ｜ result staging buffer, assigned to sDst once at the exit
    cCh      : STRING(1);   // 当前字符 [字符] ｜ current character
    sLo      : STRING(1);   // 转换后的字符 [字符] ｜ converted character
    nPos     : INT;         // 字符在码表中的位置 [索引]，1 起 ｜ character position in the code table, 1-based
    nSrcLen  : INT;         // 锁存的源文本长度 [字符]，本件唯一锁存量 ｜ latched source length, the single latched quantity
    nWritten : INT;         // 写出计数 [字符]，出口与 nSrcLen 比对 ｜ written count compared at the exit
    uCode    : UDINT;       // 码位暂存，出口单点写入 [码] ｜ code staging, written once at the exit
END_VAR
VAR CONSTANT
    DL_STL_MAXLEN : INT := 255; // 字符串上限 [字符]，与形参声明一致 ｜ string limit, matches the declarations
    DL_STL_ONE    : INT := 1;   // 单字符长度参数 [字符] ｜ single character length argument
END_VAR

// 段 1｜输出预置与残留清除：先清空再分流，拒绝路不露旧值 ｜ preset and clear before any branch, the refusal path exposes no stale value
FC_DL_StringToLowerEx := FALSE; // 预置返回失败 ｜ preset return FALSE
sDst       := '';        // 结果清空 ｜ clear the result
sTmp       := '';        // 暂存清空 ｜ clear the staging buffer
bTruncated := FALSE;     // 截断标志清零 ｜ clear the truncation flag
nKept      := 0;         // 保留计数清零 ｜ clear the kept count
nWritten   := 0;         // 写出计数清零 ｜ clear the written count
uErrorId   := 16#0000_0000; // 事件码清零 ｜ clear the event code
uCode      := 16#0000_0000; // 码位暂存清零 ｜ clear the code staging

// 段 2｜LEN 一次锁存 ｜ latch the length once
nSrcLen := LEN(sSrc);        // 源长只取一次，循环内禁重复 LEN ｜ latch the length once, never call LEN again in the loop
IF nSrcLen < 0 THEN
    nSrcLen := 0;            // 防御：异常返回值钳到零 ｜ defensive: clamp an anomalous result to zero
END_IF

// 段 3｜与上限比较，超限先置标志后分路 ｜ compare with the limit, flag first, then branch
IF nSrcLen > DL_STL_MAXLEN THEN
    bTruncated := TRUE;      // 事实先记录，早于任何写入 ｜ record the fact before any write
    IF NOT bAllowTrunc THEN
        uErrorId := 16#0001_03D4; // 故障级配对：拒绝截断以返回假表达（R45）｜ fault level, refusal expressed by FALSE
        RETURN;             // 拒绝构造，结果保持空串 ｜ refuse, result stays empty
    END_IF
    nSrcLen := DL_STL_MAXLEN; // 截断路：按上限截取 ｜ truncation path: cut to the limit
END_IF

// 段 4｜逐字符查表映射：域内转小写，域外保持并计数 ｜ per-character table mapping: convert in-domain, keep and count the rest
FOR nI := 1 TO nSrcLen DO
    cCh := MID(sSrc, DL_STL_ONE, nI);            // 位置 nI 起取一个字符 ｜ one character at position nI
    sLo := cCh;                                  // 默认保持原值 ｜ keep by default
    IF (cCh >= 'A') AND (cCh <= 'Z') THEN
        nPos := FIND('ABCDEFGHIJKLMNOPQRSTUVWXYZ', cCh);     // 大写码表定位，域内恒 1 到 26 ｜ locate in the uppercase table
        sLo  := MID('abcdefghijklmnopqrstuvwxyz', DL_STL_ONE, nPos); // 同位取小写 ｜ same position in the lowercase table
    ELSE
        nKept := nKept + DL_STL_ONE;             // 域外字符保持，累计告知 ｜ keep and count the out-of-domain char
    END_IF
    sTmp := CONCAT(sTmp, sLo);                   // 追加写出 ｜ append to the staging buffer
    nWritten := nWritten + DL_STL_ONE;           // 写出计数同步累加 ｜ sync the written count
END_FOR

// 段 5｜写出一致性校验（防御闸）：计数必须等于锁存源长 ｜ write consistency gate: the count must equal the latched length
IF nWritten <> nSrcLen THEN
    uErrorId := 16#0001_03D5;    // 故障级：写出链路异常，结果作废 ｜ fault: write chain broken, result voided
    sDst := '';                  // 结果作废清空 ｜ void and clear the result
    RETURN;                      // 返回假，bTruncated 保持已记录事实 ｜ return FALSE, the truncation fact stays recorded
END_IF

// 段 6｜出口装配：结果单点写出，码位单点写入 ｜ exit: single write for the result and the code
sDst := sTmp;                    // 暂存结果单点写出 ｜ write the staged result once
IF bTruncated THEN
    uCode := 16#0001_0499;       // 信息级：源超上限已截断 ｜ info level: source beyond the limit, truncated
END_IF
uErrorId := uCode;               // 码位单点写入 ｜ write the code once
FC_DL_StringToLowerEx := TRUE;   // 构造成功 ｜ construction succeeded
END_FUNCTION

(* ---- FC_DL_StringToUpperEx.st ---- *)
(*==============================================================================
 * 组件名称 (Component)  : FC_DL_StringToUpperEx
 * 所属子库 (Sublibrary) : DL_MathData
 * 归属目录 (Directory)  : C:\Library\DL_MathData
 * 当前版本 (Version)    : 1.0.0
 * 分类/来源标签         : 函数（FUNCTION）· 纯函数 · 字符串大写扩展转换
 *                         iec-std-wrapper / string / r37-reference
 * 兼容性   (Platform)   : CODESYS 3.5 / TwinCAT 3 / 汇川 InoProShop / 施耐德
 *                         Machine Expert；仅用 Standard.library 的 LEN / MID / CONCAT / FIND
 * 溯源声明 (Provenance) : IEC 61131-3 标准语义的道莅防御性实现——内部委托平台标准库语义，
 *                         外围统一错误码 / 钳位 / 双语注释，严禁重实现数学内核。
 * 功能一句话 (Summary)  : 把 ASCII 域内小写字母映射为大写，域外字符保持原值并计数，
 *                         全程按 R37 四步样板做长度守卫与截断分路。
 *
 * 本件存在的意义 (Why this unit exists)：
 *   各平台自带的大小写转换行为不一（有的吞掉高位字符、有的整串拒绝），本件只用
 *   标准 LEN/MID/CONCAT/FIND 做逐字符查表映射：小写字母经双码表定位转大写，
 *   其余字符原样保留并以信息码告知「有保留发生」，调用方永远知道结果里混了什么。
 *
 * 功能描述 (Function)   : 第 1 步 LEN 一次锁存源长；第 2 步与 255 上限比较；第 3 步
 *                         超限先置截断标志；第 4 步按 bAllowTrunc 分路截断写出或拒绝。
 *                         合法路径逐字符取字符：落在 'a'..'z' 域内的用 FIND 在小写
 *                         码表定位后到同位大写码表取字符，域外字符保持并累计 nKept。
 * 与既有件边界 (Boundary): 本件只做 ASCII a..z 域内映射，不做 Unicode 与本地化；
 *                         与 FC_DL_StringFixedField（改宽度不改内容）正交。
 * 码位说明 (Codes)      : 信息 16#0002_3058 存在域外字符保持原值
 *                         故障 16#0002_3059 源长度域外且未允许截断（防御闸）
 *                         故障 16#0002_305A 写出计数与源长不一致（防御校验）
 *                         段 16#02_3_58~5B 首槽信息级、次槽起故障级。
 * 依赖说明 (Depends)    : 无 DL_ 内部依赖；仅 Standard.library 的 LEN / MID / CONCAT / FIND。
 * 镜像量清单 (R38)      : nSrcLen 是本件唯一锁存量，入口一次导出，其后比较与循环
 *                         上界全部读该副本，全文不再对入参串取长度。
 * 红线自检 (Redline)    : 零全局依赖 ｜ 零 VAR_EXTERNAL ｜ 零 %I/%Q ｜ 纯 IEC 标准库
 *                         无除法故无除零面 ｜ 全变量双语同行注释 ｜ 无定时器实例
 * 修订历史 (Revision)   : 2026-11-18  v1.0.0  首版入库（R32 · 批 1）
 *============================================================================*)

FUNCTION FC_DL_StringToUpperEx : BOOL
VAR_INPUT
    sSrc        : STRING(255);      // 源文本 [ASCII]，定长 255 / Source text, fixed 255 characters
    bAllowTrunc : BOOL := FALSE;    // 允许截断，真则截断写出，假则拒绝构造 / TRUE truncates and writes, FALSE refuses
END_VAR
VAR_OUTPUT
    sDst        : STRING(255);      // 大写结果 [ASCII]，域外字符保持原值 / Uppercase result, out-of-domain chars kept
    bTruncated  : BOOL;             // 截断标志，源超上限时为真 / Set true when the source exceeded the limit
    nKept       : INT;              // 保持原值的域外字符个数 [个] / Count of kept out-of-domain characters
    uErrorId    : UDINT;            // 事件码，0 表示无事件 / Event code, zero means none
END_VAR
VAR
    sTmp     : STRING(255); // 结果累积缓冲 [ASCII]，出口一次性赋给 sDst / Result staging buffer
    cCh      : STRING(1);   // 当前字符 [字符] / Current character
    sUp      : STRING(1);   // 转换后的字符 [字符] / Converted character
    nPos     : INT;         // 字符在码表中的位置 [索引]，1 起 / Character position in the code table, 1-based
    nSrcLen  : INT;         // 锁存的源文本长度 [字符]，R38 唯一锁存量 / Latched source length, the single latched quantity
    nWritten : INT;         // 写出计数 [字符]，出口与 nSrcLen 比对 / Written count compared at the exit
    uCode    : UDINT;       // 码位暂存，出口单点写入 [码] / Code staging, written once at the exit
END_VAR
VAR CONSTANT
    DL_STU_MAXLEN : INT := 255; // 字符串上限 [字符]，与形参声明一致 / String limit, matches the declarations
    DL_STU_ONE    : INT := 1;   // 单字符长度参数 [字符] / Single character length argument
END_VAR

(* 段 1｜输出预置与残留清除：先清空再分流，拒绝路不露旧值 / Pre-set and clear before any branch *)
FC_DL_StringToUpperEx := FALSE;
sDst       := '';
sTmp       := '';
bTruncated := FALSE;
nKept      := 0;
nWritten   := 0;
uErrorId   := 16#0000_0000;
uCode      := 16#0000_0000;

(* 段 2｜R37 第 1 步：LEN 一次锁存 / Step one: latch the length once *)
nSrcLen := LEN(sSrc);
IF nSrcLen < 0 THEN
    nSrcLen := 0;                // 防御：异常返回值钳到零 / Defensive: clamp an anomalous result to zero
END_IF

(* 段 3｜R37 第 2、3 步：与上限比较，超限先置标志后分路 / Steps two and three: compare, flag, then branch *)
IF nSrcLen > DL_STU_MAXLEN THEN
    bTruncated := TRUE;          // 事实先记录，早于任何写入 / Record the fact before any write
    IF NOT bAllowTrunc THEN
        uErrorId := 16#0002_3059; // 故障级配对：本函数级故障以返回假表达（R45）/ Fault level, refusal expressed by FALSE
        RETURN;                  // 拒绝构造，结果保持空串 / Refuse, result stays empty
    END_IF
    nSrcLen := DL_STU_MAXLEN;    // 第 4 步截断路：按上限截取 / Truncation path: cut to the limit
END_IF

(* 段 4｜逐字符查表映射：域内转大写，域外保持并计数 / Per-character table mapping: convert in-domain, keep and count the rest *)
FOR nI := 1 TO nSrcLen DO
    cCh := MID(sSrc, DL_STU_ONE, nI);            // 位置 nI 起取一个字符 / One character at position nI
    sUp := cCh;                                  // 默认保持原值 / Keep by default
    IF (cCh >= 'a') AND (cCh <= 'z') THEN
        nPos := FIND('abcdefghijklmnopqrstuvwxyz', cCh);     // 小写码表定位，域内恒 1 到 26 / Locate in the lowercase table
        sUp  := MID('ABCDEFGHIJKLMNOPQRSTUVWXYZ', DL_STU_ONE, nPos); // 同位取大写 / Same position in the uppercase table
    ELSE
        nKept := nKept + DL_STU_ONE;             // 域外字符保持，累计告知 / Keep and count the out-of-domain char
    END_IF
    sTmp := CONCAT(sTmp, sUp);                   // 追加写出 / Append to the staging buffer
    nWritten := nWritten + DL_STU_ONE;           // 写出计数同步累加 / Sync the written count
END_FOR

(* 段 5｜写出一致性校验（防御闸）：计数必须等于锁存源长 / Write consistency gate: count must equal the latched length *)
IF nWritten <> nSrcLen THEN
    uErrorId := 16#0002_305A;    // 故障级：写出链路异常，结果作废 / Fault: write chain broken, result voided
    sDst := '';
    RETURN;
END_IF

(* 段 6｜出口装配：结果单点写出，码位单点写入 / Exit: single write for result and code *)
sDst := sTmp;
IF nKept > 0 THEN
    uCode := 16#0002_3058;       // 信息级：存在域外字符保持原值 / Info: out-of-domain characters kept
END_IF
uErrorId := uCode;
FC_DL_StringToUpperEx := TRUE;
END_FUNCTION

(* ---- FC_DL_StringTrim.st ---- *)
(*==============================================================================
 * 组件名称 (Component)  : FC_DL_StringTrim
 * 所属子库 (Sublibrary) : DL_MathData
 * 当前版本 (Version)    : 1.0.0
 * 兼容性   (Platform)   : CODESYS 3.5 / TwinCAT 3 / 汇川 InoProShop / Machine Expert
 *                         仅依赖 Standard.library 的标准串函数（LEN / MID）
 * 功能描述 (Function)   : 去除字符串首尾空白字符。空白集恰为四类：空格 / 制表 / 回车 /
 *                         换行，中间位置的空白原样保留（这是与"删除全部空白"的本质区别）。
 *                         双向扫描：先从头部找首个非空白位置，再从尾部找末个非空白位置，
 *                         最后一次性截取中间段，避免逐字符拼接带来的长度与性能问题。
 *                         全空白或空串输入返回空串并如实报告去除数量——这是合法结果而非错误。
 *                         扫码枪、CSV 报文、视觉结果字符串入库比对前的标准清洗步。
 * 开源溯源 (Origin)     : 原创实现。首尾裁剪为公开经典字符串处理需求；
 *                         空白字符集与位置口径依据 IEC 61131-3 标准串函数定义，
 *                         未复制任何源码。
 * 本文件内含       : FC    FC_DL_StringTrim（单 POU，无配套类型）
 * 依赖     (Depends)    : 无 DL_ 内部依赖；Standard.library: LEN / MID
 * 红线自检 (Redline)    : R1 ✓ 禁用全局存储与物理寻址 ｜ R2 ✓ 无地址直写
 *                         R3 ✓ 仅标准串函数 ｜ R4 ✓ 双循环防死锁计数 + 截取长度结构性保证
 *                         R5 ✓ 全变量中英双语同行注释 ｜ R6 N/A（纯函数，无状态机）
 *                         R7 N/A（无定时器/边沿实例）｜ R8 ✓ 长度上限与循环上限全常量化
 *
 * 【长度声明警告 / Explicit length warning（边界 B1）】
 *   输入与返回一律显式声明字符串最大长度。省略长度时平台默认上限远小于 255，
 *   超长报文会被静默截断，而截断点在运行期无任何迹象——这是串口设备集成的高频事故源。
 *
 * 【字符集边界 / Character-set boundary（边界 B2）】
 *   仅处理上述四类单字节空白。全角空格等多字节字符不属本函数职责，
 *   应在调用方做编码归一后再进入本函数。
 *
 * 【位置口径 / Position convention（边界 B3）】
 *   全程按 IEC 标准串函数口径，位置从 1 开始计数，不是从 0。
 *
 * 修订历史 (Revision)   :
 *   2026-11-14  v1.0.0  首版入库（Phase 1 第二轮 · Level 0 批次 A）
 *============================================================================*)
FUNCTION FC_DL_StringTrim : STRING(255)
VAR_INPUT
    sIn      : STRING(255);   // 原始字符串，最大 255 字符 / Source string, 255 characters max
END_VAR
VAR_OUTPUT
    bValid   : BOOL;          // 处理完整标志，FALSE = 循环保护触发 / Complete flag, FALSE = the loop guard tripped
    uTrimmed : UINT;          // 被去除的空白字符总数 [个] / Total whitespace characters removed [count]
    uErrorId : UDINT;         // 故障码，0 = 无故障 / Error code, 0 = no error
END_VAR
VAR
    nLen     : INT;           // 输入有效长度 [字符] / Effective input length [characters]
    nStart   : INT;           // 首个非空白位置（1 起始） / First non-blank position, 1-based
    nEnd     : INT;           // 末个非空白位置（1 起始） / Last non-blank position, 1-based
    nKept    : INT;           // 保留段长度 [字符] / Length of the retained segment [characters]
    sChar    : STRING(1);     // 当前检查字符 / Current character under check
    bRun     : BOOL;          // 循环继续标志 / Loop continuation flag
    nGuard   : DINT;          // 循环防死锁计数器 [次] / Loop deadlock guard counter [count]
END_VAR
VAR CONSTANT
    DL_STR_MAX_LEN  : INT  := 255;    // 串长度上限 [字符]，与类型声明一致 / Max length [characters], must match the type
    DL_STR_LOOP_MAX : DINT := 255;    // 循环防死锁上限 [次] / Loop guard limit [count]
END_VAR

(*------------------------------------------------------------------------------
 * 段 1｜结果预置（P-01 范式）：先给空串与成功标志，异常路径也必有确定返回值
 *      Safe preset: an empty result and a success flag, every path returns something
 *-----------------------------------------------------------------------------*)
FC_DL_StringTrim := '';
bValid   := TRUE;
uErrorId := 16#0000_0000;
uTrimmed := UINT#0;
nKept    := 0;

(*------------------------------------------------------------------------------
 * 段 2｜有效长度（边界 B1）：先钳位再用，后续所有位置判断都基于这一个值
 *      Effective length: clamped once and reused by every position test
 *-----------------------------------------------------------------------------*)
nLen := LEN(sIn);

IF nLen > DL_STR_MAX_LEN THEN
    nLen := DL_STR_MAX_LEN;
ELSIF nLen < 0 THEN
    nLen := 0;
END_IF

nStart := 1;
nEnd   := nLen;

(*------------------------------------------------------------------------------
 * 段 3｜头部扫描（边界 B4）：四类空白逐一比较，循环带防死锁计数
 *      Head scan: four whitespace classes compared one by one, with a loop guard
 *      全空白时 nStart 会越过 nLen，由段 5 的区间判据自然得到空串结果
 *      On an all-blank input nStart passes nLen, stage 5 then yields an empty result
 *-----------------------------------------------------------------------------*)
bRun   := (nLen > 0);
nGuard := 0;

WHILE bRun DO

    sChar := MID(sIn, 1, nStart);

    IF (sChar = ' ') OR (sChar = '$09') OR (sChar = '$0D') OR (sChar = '$0A') THEN
        nStart := nStart + 1;
        IF nStart > nLen THEN
            bRun := FALSE;
        END_IF
    ELSE
        bRun := FALSE;
    END_IF

    (* 防死锁：位置必然单调递增，仍设上限兜底，防止平台串函数异常导致位置不前进 *)
    (* Deadlock guard: the position always advances, the cap is a second line of defence *)
    nGuard := nGuard + 1;
    IF nGuard > DL_STR_LOOP_MAX THEN
        bRun     := FALSE;
        bValid   := FALSE;
        uErrorId := 16#0001_0004;
    END_IF

END_WHILE;

(*------------------------------------------------------------------------------
 * 段 4｜尾部扫描（边界 B4）：从末位向前，遇到非空白即停
 *      Tail scan: walk backwards and stop at the first non-blank
 *-----------------------------------------------------------------------------*)
IF (nStart <= nLen) AND (nEnd >= nStart) THEN

    bRun   := TRUE;
    nGuard := 0;

    WHILE bRun DO

        sChar := MID(sIn, 1, nEnd);

        IF (sChar = ' ') OR (sChar = '$09') OR (sChar = '$0D') OR (sChar = '$0A') THEN
            nEnd := nEnd - 1;
            IF nEnd < nStart THEN
                bRun := FALSE;
            END_IF
        ELSE
            bRun := FALSE;
        END_IF

        nGuard := nGuard + 1;
        IF nGuard > DL_STR_LOOP_MAX THEN
            bRun     := FALSE;
            bValid   := FALSE;
            uErrorId := 16#0001_0004;
        END_IF

    END_WHILE;

END_IF

(*------------------------------------------------------------------------------
 * 段 5｜截取（边界 B5/B6）：区间判据成立才调 MID，长度为 0 直接返回空串
 *      Extraction: MID is called only when the interval is valid, zero length returns empty
 *      区间判据是结构性保证（头部扫描保证 nStart 是首个非空白、尾部扫描保证 nEnd
 *      是末个非空白），此处再断言一次属于双保险，不承担主要防御职责
 *      The interval is structurally guaranteed; this assertion is a second line of defence
 *-----------------------------------------------------------------------------*)
IF (nStart >= 1) AND (nStart <= nLen) AND (nEnd >= nStart) AND (nEnd <= nLen) THEN

    nKept := nEnd - nStart + 1;

    IF nKept > 0 THEN
        FC_DL_StringTrim := MID(sIn, nKept, nStart);
    END_IF

ELSE
    (* 空串或全空白：合法的空结果，不是错误（边界 B5） *)
    (* Empty or all-blank input: a legal empty result, not an error *)
    nKept := 0;
END_IF

(*------------------------------------------------------------------------------
 * 段 6｜去除计数：原始有效长度减去保留长度，覆盖全部路径且不会为负
 *      Removed count: original length minus retained length, never negative
 *-----------------------------------------------------------------------------*)
IF nKept < 0 THEN
    nKept := 0;
END_IF

IF nLen >= nKept THEN
    uTrimmed := INT_TO_UINT(nLen - nKept);
ELSE
    uTrimmed := UINT#0;
END_IF
END_FUNCTION

(* ---- FC_DL_StrToHex.st ---- *)
(*
  ==================================================================
  组件名 Component  : FC_DL_StrToHex
  分类   Category   : DL_MathData
  前缀   Naming     : FC_DL_ ｜ b/n/u/f/s/a 类型前缀制（R265）
  版本   Version    : 1.0.0
  功能   Purpose    : HEX 文本 → 字节串（FC_DL_HexToStr 逆变换）：两位/
                      字节、无分隔符、接受大写与小写。解析前先过奇数长
                      度闸（LEN 奇数 → 码 02）与输出容量闸（字节预算 >
                      输出数组长度 → 码 03，不写部分数据）；逐字符经 MID
                      取样后按 '0'..'9'/'A'..'F'/'a'..'f' 判别，非法字符
                      → 码 01，三者均不写部分输出（原子性：失败即零写入）。
                      返回值 = 实际写出字节数（名实双出口）。溯源：本件
                      为「IEC 61131-3 标准语义的道莅防御性实现」，字符
                      串访问内核委托标准库函数（LEN/MID），严禁重实现内
                      核；半字节判别为纯 IEC 字面比较，非内核重实现。
  来源   Source     : iec-std-wrapper（T0-6）：IEC 61131-3 标准语义的
                      道莅防御性实现，内核委托标准库字符串函数，零内核
                      重实现
  互引   Cross-ref  : FC_DL_HexToStr（同族正变换件：字节串 → HEX 文本，
                      二者成对使用需同参数约定：大写两位/字节、无分隔符）
  平台   Platform   : 纯 IEC 61131-3（标准库字符串函数 + SHL/OR），三平台通用
  依赖   Depends    : 无 DL_ 内部依赖；标准字符串函数 LEN/MID
  红线   Redline    : R1 零全局/VAR_EXTERNAL/R2 零 %I/%Q/R3 纯 IEC 标准
                      R4 奇长闸/容量闸/非法字符闸三面显式 + 原子性零写
                      入 + 输出下标界已证（预算 ≤ 容量）/R5 全变量双语
                      同行注释/R6 纯函数无状态机（CASE 不适用）/R7 无定
                      时器与沿检测/R8 码位与界常量化
  错误码 Codes      : 01【失效级】非法字符（非 0-9/A-F/a-f），零写入
                      02【失效级】奇数长度（HEX 文本须偶数长），零写入
                      03【失效级】输出容量不足（2 字节预算 > 输出数组
                      长度），零写入
  码位反证 Note     : 01/02/03 分立依据（R90）：01 在字符面、02 在长度
                      面、03 在容量面可观测，修复入口不同（改数据/补一
                      位/扩数组）；03 若并入 01，则「扩容即可解」与「改
                      数据才能解」不可区分，故必须分立。
  验收   Acceptance : V1 '0AFF' → [0x0A,0xFF] ｜ V2 '0aff' → 同 V1（小
                      写接受）｜ V3 '0AF'（奇长）→ 码 02 ｜ V4 '0AG0'
                      → 码 01 ｜ V5 长文本/小数组 → 码 03 ｜ V6 返回值
                      = 实际字节数 = LEN/2
  变更   Revision   : 2026-11-22  v1.0.0  R67 首版（编码阶段批 3 序 1）
  ==================================================================
*)
FUNCTION FC_DL_StrToHex : UDINT
VAR_INPUT
    sHexIn : STRING(255);       // 输入 HEX 文本（两位/字节，无分隔符）/ the input hex text
END_VAR
VAR_IN_OUT
    aBytesOut : ARRAY[*] OF BYTE;  // 输出字节串（容量即数组长度）[字节] / the output byte array
END_VAR
VAR_OUTPUT
    uBytesOut : UDINT;          // 实际写出字节数 [字节]（与返回值同源，名实双出口）/ the written byte count
    bValid    : BOOL;           // 输出可用标志 [-] / the output usable flag
    nErrId    : UDINT;          // 错误码，0=正常，01/02/03 见头注 [码] / the error code [code]
END_VAR
VAR
    nChars  : UDINT;            // 输入字符数 [字符] / the input char count
    uCap    : UDINT;            // 输出数组容量 [字节] / the output array capacity
    i       : UDINT;            // 字符对遍历循环变量 / the char pair loop index
    j       : UDINT;            // 输出字节下标 / the output byte index
    k       : UDINT;            // 查表序号循环变量 / the table lookup loop index
    sHi     : STRING(1);        // 高位字符工作寄存器 / the high char register
    sLo     : STRING(1);        // 低位字符工作寄存器 / the low char register
    uHi     : BYTE;             // 高半字节值 [半字节] / the high nibble value
    uLo     : BYTE;             // 低半字节值 [半字节] / the low nibble value
    sHexTab   : STRING := '0123456789ABCDEF'; // 大写查表 [表] / the uppercase lookup table
    sHexTabLo : STRING := 'abcdef';             // 小写查表 [表] / the lowercase lookup table
END_VAR
VAR CONSTANT
    S2H_ERR_NONE  : UDINT := 16#0000_0000;  // 无错误 [码] / no error [code]
    S2H_ERR_CHR   : UDINT := 16#0000_0001;  // 码 01：非法字符 / code 01, illegal char
    S2H_ERR_ODD   : UDINT := 16#0000_0002;  // 码 02：奇数长度 / code 02, odd length
    S2H_ERR_CAP   : UDINT := 16#0000_0003;  // 码 03：输出容量不足 / code 03, capacity short
END_VAR

// 段 1｜输出预置 / segment 1, preset the outputs
uBytesOut := UDINT#0;         // 预置零写入 / preset zero written
bValid := FALSE;              // 预置不可用 / preset unusable
nErrId := S2H_ERR_NONE;       // 预置无错误 / preset no error

// 段 2｜奇数长度闸（码 02）：长度面缺陷 / segment 2, the odd length gate
nChars := LEN(sHexIn);        // 输入字符数（LEN 不含终结符）/ the char count
IF (nChars MOD 2) = UDINT#1 THEN
    nErrId := S2H_ERR_ODD;    // 奇长（补一位方可解）/ the odd length
    RETURN;
END_IF

// 段 3｜输出容量闸（码 03）：容量面缺陷，预算 = nChars/2 字节
//      segment 3, the capacity gate, the budget is nChars over two bytes
IF UPPER_BOUND(aBytesOut, 1) >= 0 THEN
    uCap := DINT_TO_UDINT(1 + UPPER_BOUND(aBytesOut, 1) - LOWER_BOUND(aBytesOut, 1));  // 数组容量 / the array capacity
ELSE
    uCap := UDINT#0;
END_IF
IF (nChars / 2) > uCap THEN
    nErrId := S2H_ERR_CAP;    // 容量不足（扩数组方可解）/ the capacity short
    RETURN;
END_IF

// 段 4｜逐对解析（委托内核：MID 取样 + 查表比较判别；下标界已证：j < nChars/2 ≤ uCap）
//      判别采用查表而非 STRING_TO_BYTE 数值转换（后者按十进制串解析，
//      字母字符不可用），表访问仍走标准 MID 内核
//      segment 4, the per pair parse, the kernel delegated to MID and table compares
FOR i := UDINT#1 TO nChars BY 2 DO        // 字符位从 1 起（MID 1 起位）/ the char position from one
    j := (i - UDINT#1) / 2;               // 输出字节下标 / the output byte index
    sHi := MID(sHexIn, 1, i);             // 高位字符 / the high char
    sLo := MID(sHexIn, 1, i + UDINT#1);   // 低位字符 / the low char
    uHi := 16#FF;                         // 非法哨兵预置（0..15 均合法，FF 不可撞）/ the illegal sentinel
    uLo := 16#FF;                         // 同上 / the same
    FOR k := UDINT#1 TO UDINT#16 DO       // 大写表查值 / the uppercase table lookup
        IF MID(sHexTab, 1, k) = sHi THEN
            uHi := UDINT_TO_BYTE(k - UDINT#1);   // 表序即半字节值 / the table order is the nibble value
            EXIT;                       // 命中即出（标准 EXIT）/ the standard exit on hit
        END_IF
    END_FOR
    IF uHi = 16#FF THEN                   // 大写未中再查小写表 / the lowercase second chance
        FOR k := UDINT#1 TO UDINT#6 DO    // 小写表 a..f / the lowercase table
            IF MID(sHexTabLo, 1, k) = sHi THEN
                uHi := UDINT_TO_BYTE(k - UDINT#1 + UDINT#10);  // a..f → 10..15 / the lower alpha nibble
                EXIT;
            END_IF
        END_FOR
    END_IF
    FOR k := UDINT#1 TO UDINT#16 DO       // 低位同法查大写表 / the low char uppercase lookup
        IF MID(sHexTab, 1, k) = sLo THEN
            uLo := UDINT_TO_BYTE(k - UDINT#1);
            EXIT;
        END_IF
    END_FOR
    IF uLo = 16#FF THEN                   // 低位小写二查 / the low char lowercase chance
        FOR k := UDINT#1 TO UDINT#6 DO
            IF MID(sHexTabLo, 1, k) = sLo THEN
                uLo := UDINT_TO_BYTE(k - UDINT#1 + UDINT#10);
                EXIT;
            END_IF
        END_FOR
    END_IF
    IF (uHi = 16#FF) OR (uLo = 16#FF) THEN     // 非法字符闸（码 01，原子性零写入）
        nErrId := S2H_ERR_CHR;                 // 字符面失效 / the char face failure
        uBytesOut := UDINT#0;                  // 零写入（原子性）/ the atomic zero write
        RETURN;
    END_IF
    aBytesOut[j] := SHL(uHi, 4) OR uLo;        // 组装字节（移位量 4 < 位宽 8，R48 合规）/ assemble the byte
END_FOR

// 段 5｜出口映射（名实双出口：返回值 = 写出字节数）/ segment 5, the exit mapping
uBytesOut := nChars / 2;      // 写出字节数 [字节] / the written byte count
FC_DL_StrToHex := uBytesOut;  // 返回值镜像（R191）/ the return mirrors the count
bValid := TRUE;               // 输出可用 / the output is usable
END_FUNCTION

(* ---- FC_DL_SwapBytes16.st ---- *)
(*==============================================================================
 * 组件名称 (Component)  : FC_DL_SwapBytes16
 * 所属子库 (Sublibrary) : DL_MathData
 * 当前版本 (Version)    : 1.0.0
 * 兼容性   (Platform)   : CODESYS 3.5 / TwinCAT 3 / 汇川 InoProShop / Machine Expert
 *                         仅依赖 Standard.library 的 SHL / SHR / AND / OR，零厂商方言
 * 功能描述 (Function)   : 16 位字高低字节互换。低字节左移 8 位升为高字节，
 *                         高字节右移 8 位降为低字节，两者按位或合成结果。
 *                         纯函数：不修改入参、无内部状态、相同输入必得相同输出；
 *                         自逆性成立，连续调用两次还原原值。
 *                         单寄存器字节序（Profibus 从站状态字、串口仪表读数）的原子构件，
 *                         同时是 32 位四排布转换的底层原子。
 * 开源溯源 (Origin)     : 原创实现。字节序定义参照 modbus.org 公开协议说明中
 *                         "单寄存器内部为大端"的事实约定；算法为公开的移位掩码法，
 *                         未复制任何厂商私有库源码，不构成衍生作品。
 * 本文件内含       : FC    FC_DL_SwapBytes16（单 POU，无配套类型）
 * 依赖     (Depends)    : 无 DL_ 内部依赖；Standard.library: SHL / SHR
 * 红线自检 (Redline)    : R1 ✓ 禁用全局存储与物理寻址 ｜ R2 ✓ 无地址直写
 *                         R3 ✓ 纯标准位运算，无字节访问方言 ｜ R4 N/A（无除法/数组/循环/浮点）
 *                         R5 ✓ 全变量中英双语同行注释 ｜ R6 N/A（纯函数，无状态机）
 *                         R7 N/A（无定时器/边沿实例）｜ R8 ✓ 移位量与掩码全常量化
 *
 * 【错误码豁免声明 / Error-code exemption】
 *   本函数不设 uErrorId 输出引脚。理由：16 位字节互换的全定义域均为合法输入，
 *   不存在任何运行期失败路径；恒为 0 的错误码引脚只会增加调用方噪音。
 *   沿用首轮 FC_DL_PackBitsToWord 的显式豁免先例（ROUND_PLAN_R2 §2.8 决策 P3）。
 *
 * 【实现选择 / Implementation choice】
 *   仅用移位 + 掩码 + 按位或，禁止任何按字节访问的厂商方言语法（R3 关键考点）。
 *   移位量经 VAR CONSTANT 统一给出，避免字面量散落造成口径漂移。
 *
 * 修订历史 (Revision)   :
 *   2026-11-14  v1.0.0  首版入库（Phase 1 第二轮 · Level 0 批次 A）
 *============================================================================*)
FUNCTION FC_DL_SwapBytes16 : WORD
VAR_INPUT
    uValue : WORD;                       // 原始 16 位字 / Source word
END_VAR
VAR
    uLow   : WORD;                       // 低字节缓存（左移后成为高字节）/ Low byte buffer, shifted up to the high byte
    uHigh  : WORD;                       // 高字节缓存（右移后成为低字节）/ High byte buffer, shifted down to the low byte
END_VAR
VAR CONSTANT
    DL_SWAP_SHIFT8 : UDINT := 8;         // 字节移位量 [bit]，全库统一口径 / Byte shift width [bit], unified library-wide
    DL_MASK_LOW8   : WORD := 16#00FF;    // 低 8 位掩码 / Low-byte mask
END_VAR

(*------------------------------------------------------------------------------
 * 段 1｜安全预置（P-01 范式）：任何异常路径返回原值，绝不返回 0
 *      Safe preset: every exceptional path returns the source value, never zero
 *-----------------------------------------------------------------------------*)
FC_DL_SwapBytes16 := uValue;

(*------------------------------------------------------------------------------
 * 段 2｜字节分离与重装（边界 B1/B5）：全程在 WORD 域内运算，无跨类型转换
 *      Byte separation and reassembly: WORD domain only, no cross-type conversion
 *      低位字节左移 8 位升为高位，高位字节右移 8 位降为低位，再按位或合成
 *      Low byte shifts up by 8, high byte shifts down by 8, then bitwise OR
 *-----------------------------------------------------------------------------*)
uLow  := SHL(uValue AND DL_MASK_LOW8, DL_SWAP_SHIFT8);
uHigh := SHR(uValue, DL_SWAP_SHIFT8);

(*------------------------------------------------------------------------------
 * 段 3｜结果回写（边界 B4）：纯函数出口唯一，无副作用
 *      Result write-back: single exit, no side effect
 *      验收向量：16#1A2B → 16#2B1A；自逆性 Swap(Swap(x)) = x 对全字域成立
 *      Acceptance vector: 16#1A2B -> 16#2B1A; self-inverse over the whole word domain
 *-----------------------------------------------------------------------------*)
FC_DL_SwapBytes16 := uLow OR uHigh;
END_FUNCTION

(* ---- FC_DL_SwapBytes64.st ---- *)
(*
    FC_DL_SwapBytes64 —— LWORD 全字节逆序
    ------------------------------------------------------------------
    分类      : DL_MathData / Convert
    前缀      : FC_DL_
    版本      : 1.0.0
    溯源      : IEC 61131-3 标准语义的道莅防御性实现（LWORD 8 字节全逆序）；
                拆合本件自有的移位与掩码，字节逆序委托库内既有件 FC_DL_SwapBytes32
                （同库资产复用，R12 PortDiagBoard 先例），不重实现字节序内核；
                掩码常量、拆合顺序与码位 100% 自有；
                clean-room 重写，未复制任何闭源厂商源码，参考实现仅限 MIT/Apache 许可
    平台      : 纯 IEC 61131-3，CODESYS V3.5+ / TwinCAT 3 / InoProShop 通用
    作者      : 道莅代码库 · PLC编程专家（R20）
    ------------------------------------------------------------------
    功能说明  : EtherCAT / CANopen 伺服与智能仪表的 64 位累计量（绝对编码器位置、
                累计流量、电表总电量）按小端直出时，进 PLC 后必须做全字节逆序才与
                上位机的显示口径一致。字节序族已有 16 位与 32 位件，64 位一直是缺口。
                核心防御：① 移位量恒为 32，结构性小于 LWORD 位宽 64，
                   禁出现 SHL/SHR(x, 位宽) 这类跨平台未定义写法（R48 纪律）；
                ② 拆高低 32 位后各自委托 FC_DL_SwapBytes32 做四字节全反序，
                   再把低位的反序结果放到高位、高位反序结果放低位——
                   全字节逆序在 64 位域上等价于「两个 32 位各自逆序再交换半区」；
                ③ 掩码 16#0000_0000_FFFF_FFFF 全常量化，禁裸值；
                ④ 本件是全域双射：任何 LWORD 输入都有唯一确定的输出，不存在非法输入，
                   故信息槽与故障槽按规格全预留禁用，也不为「不存在的错误」虚构码位；
                ⑤ 多次调用幂等：逆序两次即还原，验收向量见下。
                验收向量：输入 16#0102_0304_0506_0708 输出 16#0807_0605_0403_0201。
                职责边界：16 位逆序归 FC_DL_SwapBytes16，32 位四排布归一归 FC_DL_SwapBytes32；
                本件只管 64 位全字节逆序。
    编译门槛  : 主路径依赖平台内建 SHL / SHR（ANY_BIT 语义）、LWORD_TO_DWORD、DWORD_TO_LWORD，
                以及 Standard.library 的位串函数，三平台标准库均提供。
                依赖库内 FC_DL_SwapBytes32 与其配套枚举 E_DL_ByteOrder（同子库，编译顺序无要求）。
    错误码    : 16#0001_0424 预留禁用（信息级，不得挪用——全双射无信息出口）
                16#0001_0425 预留禁用（信息级，不得挪用）
                16#0001_0354 预留禁用（故障级，不得挪用——全域双射不存在非法输入）
                16#0001_0355 预留禁用（故障级，不得挪用）
                16#0001_0356 预留禁用（故障级，不得挪用）
    码位总账  : 16#0001_0424 预留 / 16#0001_0425 预留 ｜ 16#0001_0354 预留 / 16#0001_0355 预留 / 16#0001_0356 预留
    状态机    : R6 标注 N/A —— 本组件为纯函数无顺序状态机，无 CASE 可写，非法状态不可能出现
    采样约定  : 本件无定时器、无沿检测、无状态；单拍纯计算，结论与任务周期无关。
    修订记录  : 2026-11-16 v1.0.0 首次入库（R20）
*)
FUNCTION FC_DL_SwapBytes64 : LWORD
VAR_INPUT
    liIn             : LWORD;                 // 输入值 [位图]，全域 0~2^64−1 / input value [bitmap], full LWORD domain
END_VAR
VAR_OUTPUT
    eErr             : UDINT;                 // 错误码，0=正常（本件恒 0，五槽全预留）/ error id, always 0 here as all five slots are reserved
    bError           : BOOL;                  // 故障标志，本件恒 FALSE / error flag, always FALSE here
    bValid           : BOOL;                  // 返回值是否可用，本件恒 TRUE / return usable, always TRUE here
END_VAR
VAR CONSTANT
    DL_SHIFT_DWORD   : UINT := 32;            // 半区移位量 [bit]，结构性小于位宽 64 / half word shift [bit], structurally below the width of 64
    DL_MASK_LO32     : LWORD := 16#0000_0000_FFFF_FFFF; // 低 32 位掩码 [位图] / mask of the low 32 bits [bitmap]
    DL_LWORD_ZERO    : LWORD := 16#0000_0000_0000_0000;  // 长字零常量，避免裸字面量 [位图] / long word zero constant [bitmap]
END_VAR
VAR
    uDwHi            : DWORD;                 // 高 32 位半区 [位图] / the high 32-bit half [bitmap]
    uDwLo            : DWORD;                 // 低 32 位半区 [位图] / the low 32-bit half [bitmap]
    uDwHiRev         : DWORD;                 // 高半区四字节逆序结果 [位图] / byte reversed high half [bitmap]
    uDwLoRev         : DWORD;                 // 低半区四字节逆序结果 [位图] / byte reversed low half [bitmap]
    liOut            : LWORD;                 // 合成结果中间量 [位图] / composed result intermediate [bitmap]
END_VAR

// 段 1｜返回值与错误状态预置 / segment 1, preset return value and error status
FC_DL_SwapBytes64 := DL_LWORD_ZERO;           // 缺省返回全零 [位图] / default returns all zero [bitmap]
eErr := 0;                                    // 五槽全预留，恒无错误 / all five slots are reserved, no error is ever raised
bError := FALSE;                              // 本件无故障出口 / no fault exit exists
bValid := FALSE;                              // 预置不可用，段 5 置位 / preset invalid, set TRUE in stage 5
liOut := DL_LWORD_ZERO;                       // 合成中间量清零 / clear the composition intermediate

// 段 2｜拆半区：移位量 32 恒小于位宽 64，掩码全常量化 / segment 2, split the halves safely
uDwHi := LWORD_TO_DWORD(SHR(liIn, DL_SHIFT_DWORD));      // 右移半区宽取高 32 位 [位图] / shift by the half width to take the high 32 bits [bitmap]
uDwLo := LWORD_TO_DWORD(liIn AND DL_MASK_LO32);          // 掩码取低 32 位 [位图] / mask the low 32 bits [bitmap]

// 段 3｜半区各自委托库内既有件做四字节全反序（不重实现字节序内核）/ segment 3, delegate each half to the existing library component
uDwHiRev := FC_DL_SwapBytes32(uRaw := uDwHi, eRawOrder := eDcba); // 高半区全反序 [位图] / byte reverse of the high half [bitmap]
uDwLoRev := FC_DL_SwapBytes32(uRaw := uDwLo, eRawOrder := eDcba); // 低半区全反序 [位图] / byte reverse of the low half [bitmap]

// 段 4｜合成：低半区反序结果进高 32 位，高半区反序结果进低 32 位 / segment 4, compose the reversed halves
liOut := SHL(DWORD_TO_LWORD(uDwLoRev), DL_SHIFT_DWORD) OR DWORD_TO_LWORD(uDwHiRev); // 全字节逆序结果 [位图] / the full byte reversed result [bitmap]

// 段 5｜发布结果 / segment 5, publish the result
FC_DL_SwapBytes64 := liOut;                   // 输出全字节逆序值 [位图] / publish the byte reversed value [bitmap]
bValid := TRUE;                               // 全域双射恒可用 / a total bijection is always usable
bError := FALSE;                              // 无故障出口（双保险）/ no fault exit exists, second line of defence
END_FUNCTION

(* ---- FC_DL_TanDegChk.st ---- *)
(*==============================================================================
 * 名称 : FC_DL_TanDegChk —— 角度制正切（含 |cos| 不可定义防护）
 * 分类 / 前缀 / 版本 : DL_MathData / FC_DL_ / 1.0.0
 * 溯源 : 开源语义参考（OSCAT/AixOCAT 族，MIT）或 clean-room IEC 实现，未复制源码
 * 平台 : 纯 IEC 61131-3
 * 功能说明 : 返回 tan(fDeg)：内部换算弧度后先求 COS 判可定义性，|cos|<1.0E-12
 *            （90°/270° 等渐近角附近）时判不可定义，返回 0.0、bValid=FALSE
 *            并置 eErr；可定义时返回标准 TAN。
 *            边界处理：输入非有限（NaN/±Inf）或 |fDeg|>1.0E12 置 eErr 返回 0.0。
 * 错误码 : 16#0001_1B0B = |cos|<1.0E-12（正切不可定义），或输入非有限 / 超安全量程 ±1.0E12
 *          eErr=0 且 bValid=TRUE 表示返回值可用
 * 状态机 : R6 标注 N/A（纯函数无顺序状态，以本节替代 ELSE 兜底）
 * 红线 : R1/R2/R3 ✓ 零全局/零IO/纯IEC ｜ R4 ✓ 非有限拦截/除零防护（渐近角）/量程防护 ｜ R10 ✓ 标准转换 ｜ R11 ✓ 分号收尾 ｜ R15 ✓ 无保留字撞名
 * 修订记录 : 2026-11-23 v1.0.0 首次入库（R76）
 *============================================================================*)
FUNCTION FC_DL_TanDegChk : LREAL
VAR_INPUT
    fDeg : LREAL;    // 输入角 [度] / input angle in degrees
END_VAR
VAR_OUTPUT
    eErr   : UDINT;    // 故障码，0=正常，1B0B=不可定义或非有限 / error code
    bError : BOOL;     // TRUE=本件发生故障 / TRUE when fault occurred
    bValid : BOOL;     // TRUE=返回值可用 / TRUE when return value is usable
END_VAR
VAR
    _fRad : LREAL;     // 换算后的弧度角 [rad] / converted angle in radians
    _fCos : LREAL;     // 余弦值（可定义性判据）/ cosine value used as guard
END_VAR

FC_DL_TanDegChk := 0.0;                      // 返回值预设 0.0 / preset return to zero
eErr   := 16#0000_0000;                      // 故障码清零 / clear error code
bError := FALSE;                             // 故障标志清零 / clear error flag
bValid := TRUE;                              // 预设输出可用 / preset valid flag

IF (fDeg <> fDeg) OR ((fDeg - fDeg) <> (fDeg - fDeg))    // NaN 或 ±Inf / NaN or infinite
   OR (ABS(fDeg) > 1.0E12) THEN              // 超安全量程 / beyond safe range
    eErr   := 16#0001_1B0B;                  // 置故障码 / set error code
    bError := TRUE;                          // 置故障标志 / set error flag
    bValid := FALSE;                         // 返回值不可用 / return not usable
    RETURN;                                  // 返回 0.0 / return zero
END_IF

_fRad := fDeg * 3.14159265358979323846 / 180.0;    // 度转弧度 / degrees to radians
_fCos := COS(_fRad);                         // 求余弦作渐近防护判据 / cosine as asymptote guard

IF ABS(_fCos) < 1.0E-12 THEN                 // 渐近角附近不可定义 / near-asymptote undefined
    eErr   := 16#0001_1B0B;                  // 置不可定义码 / set undefined code
    bError := TRUE;                          // 置故障标志 / set error flag
    bValid := FALSE;                         // 返回值不可用 / return not usable
    FC_DL_TanDegChk := 0.0;                  // 返回 0.0（契约约定）/ return zero per contract
    RETURN;                                  // 提前收口 / early exit
END_IF

FC_DL_TanDegChk := TAN(_fRad);               // 可定义域内取正切 / tangent in defined domain

END_FUNCTION

(* ---- FC_DL_TanEx.st ---- *)
(*==============================================================================
 * 组件名称 (Component)  : FC_DL_TanEx
 * 所属子库 (Sublibrary) : DL_MathData
 * 当前版本 (Version)    : 1.0.0
 * 兼容性   (Platform)   : CODESYS 3.5 / TwinCAT 3 / 汇川 InoProShop / Machine Expert
 *                         仅依赖 Standard.library 的 TAN / COS / ABS 内建函数，
 *                         不重实现三角内核，无厂商数学方言依赖
 * 功能一句话 (Summary)  : 正切防御包装：弧度制输入，π/2 + kπ 周期奇点
 *                         双闸拦截（cos 容差闸 + 幅值上限闸），委托内建 TAN。
 * 功能描述 (Function)   : 对弧度制角度 fX 求正切。三道闸门按次序写死：
 *                         ① 非有限复检先行（NaN 用 x <> x 判据、无穷用
 *                         ABS(x) 超有限性上界判据）；② π/2 极点容差闸——
 *                         用内建 COS 求 |cos(fX)|（不自写级数），|cos| <
 *                         1.0E-12 判为极点邻域，返回 0.0 + 故障码；
 *                         ③ 域内委托内建 TAN，结果做非有限与幅值双重复检：
 *                         |tan| 超过 1.0E6 幅值上限判为奇点域（内建 TAN 在
 *                         极点可能返回天文数字而非 Inf，幅值闸必须兜住）。
 * 溯源     (Origin)     : IEC 61131-3 标准语义的道莅防御性实现
 *                         （接口语义由 IEC 61131-3 定义，clean-room 重写，
 *                         参考公开标准条款）
 * 码位     (Diag Codes) : 故障级 16#0001_022A（本件独占）：
 *                           极点邻域（|cos(fX)| < 1.0E-12）、输入/输出非有限
 *                           或幅值爆炸（|tan| > 1.0E6）——三况同码，均判为
 *                           奇点域，返回安全值 0.0。
 * 类型裁定 (Type Note)  : 码位段 16#0001_xxxx 为全库共享 32 位段，WORD 容量不足，
 *                         故 eErr 采用 UDINT 承载（与库内 uErrorId : UDINT 惯例
 *                         一致，沿 R14 批 3 同一裁定）。
 * 单位声明 (Unit Note)  : 输入 fX 单位为弧度 [rad]，非角度制；角度制调用方
 *                         先乘 π/180 显式转换后再调用，本件不做隐式换算。
 * 依赖     (Depends)    : 无 DL_ 内部依赖；Standard.library: TAN / COS / ABS
 * 红线自检 (Redline)    : R1 ✓ 零全局变量与外部变量引用 ｜ R2 ✓ 零物理 IO 地址直写
 *                         R3 ✓ 纯 IEC 61131-3 ｜ R4 ✓ 三道闸门次序写死 + 双重复检
 *                         R5 ✓ 全变量中英双语同行注释
 *                         R6 N/A（纯函数，无 CASE/ENUM 状态机，按批 4 口径标 N/A）
 *                         R7 N/A（FC 为纯函数，无实例调用，头注释显式说明）
 * 防御行为声明 (Defense): ① 弧度制输入 [rad]，不做隐式角度换算（单位声明节）；
 *                         ② 非有限复检先行：NaN 判据 fX <> fX（NaN 与任何值
 *                           包括自身比较均为不等，库内既有写法）、无穷判据
 *                           ABS(fX) > 1.0E308，命中即不调内建、早退返回 0.0；
 *                         ③ 极点容差闸前置：|cos(fX)| < 1.0E-12 判为 π/2 + kπ
 *                           周期奇点邻域，cos 由内建求（严禁自写泰勒级数），
 *                           返回 0.0 + 故障码，杜绝幅值爆炸值进入下游；
 *                         ④ 幅值上限闸兜底：内建 TAN 在极点邻域可能返回
 *                           天文数字有限值而非 Inf，|tan| > 1.0E6 判奇点域
 *                           返回 0.0 + 故障码（非有限与幅值双判据同码 022A）；
 *                         ⑤ 1.0E-12 容差与 1.0E6 幅值上限、1.0E308 有限性
 *                           上界均提为只读常量，禁魔法数；
 *                         ⑥ 浮点全程不用等号直比判数值相等，仅用 < > 与
 *                           NaN 自不等判据，符合浮点容差红线口径。
 * 修订历史 (Revision)   :
 *   2026-11-16  v1.0.0  首版入库（R14 批 4 · T0 快车道）
 *============================================================================*)
FUNCTION FC_DL_TanEx : LREAL
VAR_INPUT
    fX : LREAL; // 自变量 [rad]，弧度制，非角度制 / Argument [rad], radians, not degrees
END_VAR
VAR_OUTPUT
    eErr : UDINT; // 错误码，16#0001_022A=极点邻域/非有限/幅值爆炸（奇点域），0=无事件 / Error code, 16#0001_022A=pole neighborhood or non-finite or amplitude blow-up (singular domain), 0=no event
END_VAR
VAR CONSTANT
    DL_TAN_FINITE : LREAL := 1.0E308; // 有限性上界 [无量纲]，超界判无穷（库内既有写法）/ Finiteness bound, values beyond treated as infinity (library idiom)
    DL_TAN_EPS    : LREAL := 1.0E-12; // 极点容差 [无量纲]，|cos| 低于此判奇点邻域 / Pole tolerance, |cos| below this means pole neighborhood
    DL_TAN_SAT    : LREAL := 1.0E6;   // 幅值上限 [无量纲]，|tan| 超此判奇点域 / Amplitude ceiling, |tan| above this means singular domain
END_VAR

(*------------------------------------------------------------------------------
 * 段 1｜返回值与错误码预置：先归零，任何早退路径都不会留下脏码
 *      Preset return value and error code so no early-exit path leaves a stale code
 *-----------------------------------------------------------------------------*)
FC_DL_TanEx := 0.0;   // 返回值预置 0.0（安全值，绝不输出 NaN / 天文数字）/ Preset return to 0.0 (safe value, never NaN or astronomical value)
eErr        := 16#0000_0000;   // 错误码预置无事件 / Preset error code to no event

(*------------------------------------------------------------------------------
 * 段 2｜闸门一：非有限复检先行（防御声明②），NaN / 无穷不进内建内核
 *      Gate 1: non-finite recheck first (defense note 2), NaN and infinity
 *      never reach the built-in kernel
 *-----------------------------------------------------------------------------*)
IF (fX <> fX) OR (ABS(fX) > DL_TAN_FINITE) THEN
    eErr := 16#0001_022A;   // 故障码：输入非有限，判奇点域，拦截早退 / Fault: non-finite input, singular domain, intercepted
    RETURN;                 // 返回预置安全值 0.0 / Return preset safe value 0.0
END_IF

(*------------------------------------------------------------------------------
 * 段 3｜闸门二：π/2 极点容差闸前置（防御声明③）——|cos(fX)| < 1.0E-12
 *      判为周期奇点 π/2 + kπ 邻域，cos 委托内建求，不自写级数
 *      Gate 2: pole tolerance gate ahead (defense note 3) — |cos(fX)| below
 *      1.0E-12 means the periodic singularity neighborhood; cos via the
 *      built-in, never a hand-rolled series
 *-----------------------------------------------------------------------------*)
IF ABS(COS(fX)) < DL_TAN_EPS THEN
    eErr := 16#0001_022A;   // 故障码：极点邻域（π/2 + kπ），返回安全值 0.0 / Fault: pole neighborhood (pi/2 + k*pi), safe value 0.0 returned
    RETURN;                 // 返回预置安全值 0.0 / Return preset safe value 0.0
END_IF

(*------------------------------------------------------------------------------
 * 段 4｜域内委托内建内核（防御声明①④）：极点邻域外委托内建 TAN
 *      In-domain delegation to the built-in kernel (defense notes 1 and 4):
 *      outside the pole neighborhood, delegate to the built-in TAN
 *-----------------------------------------------------------------------------*)
FC_DL_TanEx := TAN(fX);   // 委托内建 TAN 内核，不自实现三角 / Delegate to the built-in TAN kernel, no re-implementation

(*------------------------------------------------------------------------------
 * 段 5｜闸门三：结果双重复检（防御声明④⑤）——非有限或 |tan| 超 1.0E6
 *      幅值上限均判奇点域，兜住「极点返回天文数字而非 Inf」的平台差异
 *      Gate 3: dual result recheck (defense notes 4 and 5) — non-finite or
 *      |tan| above the amplitude ceiling both mean singular domain, catching
 *      platforms that return huge finite values instead of Inf at poles
 *-----------------------------------------------------------------------------*)
IF (FC_DL_TanEx <> FC_DL_TanEx) OR (ABS(FC_DL_TanEx) > DL_TAN_FINITE) OR (ABS(FC_DL_TanEx) > DL_TAN_SAT) THEN
    FC_DL_TanEx := 0.0;    // 兜底安全值 0.0 / Bottom-line safe value 0.0
    eErr := 16#0001_022A;   // 故障码：输出非有限或幅值爆炸，判奇点域 / Fault: non-finite or blown-up output, singular domain
END_IF
END_FUNCTION

(* ---- FC_DL_ThdCalc.st ---- *)
(*
  ==================================================================
  组件名 Component  : FC_DL_ThdCalc
  分类   Category   : DL_MathData
  复杂度 Complexity  : 低
  版本   Version    : 1.0.0
  功能   Purpose    : 总谐波失真率 THD = √(Σ h₂..hN²) / |h₁|。输入为幅值序列
                      （0 号位基波，1..N-1 为各次谐波），基波近零或非有限立即
                      置码并拒绝相除，谐波幅值按绝对值域参与（幅值约定）。
  来源   Source     : self-std（IEC 61131-3 标准数学语义自研聚合层）
  溯源   Origin     : THD 定义属公开电能质量语义，道莅 clean-room 自研实现，
                      未复制任何厂商私有库源码。
  平台   Platform   : 纯 IEC 61131-3（SQRT / ABS / FOR），三平台通用
  分工声明 Split     : 与 FC_DL_HarmonicSpectrumBin（频点分箱属主）与
                      FC_DL_FftRadix2（变换属主）分工——本件只做幅值序列的
                      聚合比值，不分箱、不做变换、不判谐波次数合法性。
  作者   Author     : 道莅代码库 · PLC 编程专家（R60）
  ------------------------------------------------------------------
  边界 Boundary     :
                      一 基波判据：|h₁| < 1E-9 判不可算，置故障级码并返回 0，
                         全程不执行除法（除零前置拦截）；
                      二 非有限判据：基波与参与谐波逐个用 x <> x（NaN）与
                         (x−x) <> (x−x)（Inf）双判，命中即三件套置位（R258）；
                      三 幅值域约定：谐波幅值取绝对值参与平方和，负幅值视为
                         相位翻转的幅值等价（本函数只出比值，不保留符号）；
                      四 计数钳位 [2, 元素容量]：少于 2 个元素无谐波可算，置
                         信息级码并返回 0；超容量钳位续算并置同一信息级码；
                      五 只读输入数组，不改调用方数据。
  错误码   Codes    :
    16#0001_0623【信息级】谐波计数越域已钳位（<2 或 >64）
    16#0001_0624【故障级】基波幅值近零（< 1E-9），THD 不可算
    16#0001_0625【故障级】样本含非有限值，THD 不可算
  验收   Acceptance :
    算法已证（脚本）：未跑 ｜ 编译器已证（三平台）：未跑
    V1 h = 100 / 10 / 10，个数 3 → THD = 0.141421（√200/100）
    V2 h = 100 / 0，个数 2 → THD = 0.0，bValid = TRUE
    V3 h₁ = 0 → 码 0624、bValid = FALSE、fThd = 0
    V4 h₂ = NaN → 码 0625、bValid = FALSE、fThd = 0
  修订记录 Revision  :
    2026-11-21  v1.0.0  R60 首版（批 2 · 序号 7）
  ==================================================================
*)
FUNCTION FC_DL_ThdCalc : LREAL
VAR_IN_OUT
    afHarm : ARRAY[0..63] OF LREAL; // 幅值序列 [幅值]，0 号位基波 / the amplitude series with the fundamental at the entry zero
END_VAR
VAR_INPUT
    nCount : DINT; // 幅值元素数（含基波）[个]，合法域 2..64 / the element count including the fundamental, legal from two to sixty four
END_VAR
VAR_OUTPUT
    bValid : BOOL;  // 结果可用标志 [-] / the result usable flag
    eErr   : UDINT; // 错误码，0 = 正常 / the error code, zero is ok
    bError : BOOL;  // 错误标志，eErr 非 0 时为真 / the error flag, true when eErr is nonzero
    nUsed  : DINT;  // 实际参与元素数 [个] / the element count actually used
END_VAR
VAR
    nI      : DINT;  // 遍历索引 [个] / the loop index
    fBase   : LREAL; // 基波幅值绝对值 [幅值] / the absolute fundamental amplitude
    fSqSum  : LREAL; // 谐波平方和 [幅值平方] / the harmonic square sum
    fV      : LREAL; // 当前谐波幅值工作副本 [幅值] / the current harmonic amplitude copy
    bNonFin : BOOL; // 非有限命中标志 [-] / the non finite hit flag
    bClamp  : BOOL; // 计数钳位标记 [-] / the count clamp flag
END_VAR
VAR CONSTANT
    DL_THD_NMAX   : DINT := 64;    // 元素容量上界 [个]，与数组容量一致 / the element capacity aligned with the array
    DL_THD_FLOOR  : LREAL := 1.0E-9; // 基波近零判据 [幅值] / the fundamental near zero criterion
END_VAR

// 段 1｜返回值与错误状态预置安全值（四段式第一段，R45）+ 局部量显式预置（R254）/ segment 1, the preset of the return, the codes and the local guards
FC_DL_ThdCalc := 0.0; // 返回值预置安全值零 / preset the return to zero
bValid := FALSE; // 有效标志预置假 / preset the validity false
eErr := 16#0000_0000; // 错误码预置正常 / preset the code to ok
bError := FALSE; // 错误标志预置假 / preset the error flag false
nUsed := 0; // 参与元素数预置零 / preset the used count zero
fBase := 0.0; // 基波幅值预置零 / preset the fundamental zero
fSqSum := 0.0; // 平方和预置零 / preset the square sum zero
fV := 0.0; // 谐波副本预置零 / preset the harmonic copy zero
bNonFin := FALSE; // 非有限标志预置假 / preset the non finite flag false
bClamp := FALSE; // 钳位标记预置假 / preset the clamp flag false

// 段 2｜计数域闸（少于 2 早退，超容量钳位，边界四）/ segment 2, the count domain gate
IF nCount < 2 THEN // 无谐波可算 / no harmonic exists
    eErr := 16#0001_0623; // 信息级：计数越域已钳位 / informational, the count clamped
    bError := TRUE; // 置错误标志（信息级随事件置位惯例）/ raise the error flag
    RETURN; // 早退：bValid 保持假、返回 0 / early return with the validity false
END_IF
nUsed := nCount; // 域内接管 / take the count inside the domain
IF nUsed > DL_THD_NMAX THEN // 超容量 / above the capacity
    nUsed := DL_THD_NMAX; // 钳到容量 / clamp to the capacity
    bClamp := TRUE; // 置钳位标记 / raise the clamp flag
    eErr := 16#0001_0623; // 信息级：计数越域已钳位 / informational, the count clamped
    bError := TRUE; // 置错误标志 / raise the error flag
END_IF

// 段 3｜基波有限性与近零闸（除零前置拦截，边界一二）/ segment 3, the fundamental finiteness and near zero gate
fBase := ABS(afHarm[0]); // 基波取绝对值（幅值域约定，边界三）/ take the absolute fundamental amplitude
IF (fBase <> fBase) OR ((fBase - fBase) <> (fBase - fBase)) THEN // 基波非有限（NaN 自反 + Inf 差值自减）/ the fundamental is not finite
    bNonFin := TRUE; // 置非有限标志 / raise the non finite flag
END_IF
IF bNonFin THEN // 非有限即拒算 / refuse the computation on a non finite value
    eErr := 16#0001_0625; // 故障级：样本含非有限值 / fault grade, a non finite sample exists
    bError := TRUE; // 置错误标志（R45 配对）/ raise the error flag, paired with the fault code
    bValid := FALSE; // 结果不可用 / the result void
    RETURN; // 早退：三件套已置（R258）/ early return with the triple raised
END_IF
IF fBase < DL_THD_FLOOR THEN // 基波近零，不可相除 / the fundamental near zero cannot divide
    eErr := 16#0001_0624; // 故障级：基波幅值近零 / fault grade, the fundamental near zero
    bError := TRUE; // 置错误标志（R45 配对）/ raise the error flag, paired with the fault code
    bValid := FALSE; // 结果不可用 / the result void
    RETURN; // 早退：全程未执行除法 / early return without any division
END_IF

// 段 4｜谐波平方和累加（逐个非有限剔除为拒算，不静默跳过）/ segment 4, the harmonic square sum with an explicit refusal
FOR nI := 1 TO nUsed - 1 DO // 有界循环（nUsed 已钳 ≤64）/ the bounded loop
    fV := ABS(afHarm[nI]); // 谐波取绝对值 / take the absolute amplitude
    IF (fV <> fV) OR ((fV - fV) <> (fV - fV)) THEN // 谐波非有限 / a non finite harmonic
        bNonFin := TRUE; // 置非有限标志 / raise the non finite flag
    ELSE // 有限谐波参与累加 / a finite harmonic participates
        fSqSum := fSqSum + fV * fV; // 平方累加 / accumulate the square
    END_IF
END_FOR
IF bNonFin THEN // 任一谐波非有限 / any harmonic is not finite
    eErr := 16#0001_0625; // 故障级：样本含非有限值 / fault grade, a non finite sample exists
    bError := TRUE; // 置错误标志（R45 配对）/ raise the error flag, paired with the fault code
    bValid := FALSE; // 结果不可用 / the result void
    FC_DL_ThdCalc := 0.0; // 返回值回安全值（不泄半结果）/ the return back to the safe zero
    RETURN; // 早退 / early return
END_IF

// 段 5｜比值计算与结果复检（除子已证 ≥ 1E-9）/ segment 5, the ratio and the result recheck
FC_DL_ThdCalc := SQRT(fSqSum) / fBase; // THD = √Σh² / |h₁|（除子已证非零）/ the ratio with a proven nonzero divisor
IF (FC_DL_ThdCalc <> FC_DL_ThdCalc) OR ((FC_DL_ThdCalc - FC_DL_ThdCalc) <> (FC_DL_ThdCalc - FC_DL_ThdCalc)) THEN // 结果非有限兜底（R258 三件套）/ the non finite result guard
    FC_DL_ThdCalc := 0.0; // 兜底安全值 / the bottom-line safe value
    eErr := 16#0001_0625; // 故障级：结果非有限（平方和溢出）/ fault grade, the non finite result
    bError := TRUE; // 置错误标志（R45 配对）/ raise the error flag, paired with the fault code
    bValid := FALSE; // 结果不可用 / the result void
ELSE // 结果有限 / a finite result
    bValid := TRUE; // 结果可用 / the result is usable
END_IF
END_FUNCTION

(* ---- FC_DL_TimeAbsSat.st ---- *)
(*
    FC_DL_TimeAbsSat —— TIME 绝对值（负 TIME 平台歧义统一口径）
    ------------------------------------------------------------------
    分类      : DL_MathData / TimeArith
    前缀      : FC_DL_
    版本      : 1.0.0
    溯源      : IEC 61131-3 标准语义的道莅防御性实现（TIME 取绝对值，含 −MAX−1 边界）；
                委托平台内建 TIME_TO_DINT / DINT_TO_TIME 完成显式换算，本件不重实现时间算术内核；
                负值口径统一、不可表边界饱和、错误分级与码位 100% 自有；
                clean-room 重写，未复制任何闭源厂商源码，参考实现仅限 MIT/Apache 许可
    平台      : 纯 IEC 61131-3，CODESYS V3.5+ / TwinCAT 3 / InoProShop 通用
    作者      : 道莅代码库 · PLC编程专家（R20）
    ------------------------------------------------------------------
    功能说明  : 偏差、超调、节拍抖动的幅值统计经常要把「正的偏差」与「负的偏差」合成同一量纲。
                但 TIME 在 IEC 61131-3 里是时长型：各平台对负 TIME 的文本解释、比较行为与
                隐式转换口径并不一致（R55 教训），直接用平台取反极易得到一个天文正数。
                本件是负 TIME 口径的原子化统一出口：任何需要幅值的场景都走它，不再就地取反。
                核心防御：① 一切判定都在 DINT 毫秒域内进行，显式 TIME_TO_DINT 取值、
                   显式 DINT_TO_TIME 回装，全程禁隐式转换；
                ② −MAX−1 案先判后算：DINT 最小值的相反数无法用 DINT 表，直接取反会静默
                   回绕成一个负数，故先判边界，再取反；
                ③ 边界判据按「极限值 → 类型可表性」反算，取严格小于 −2147483647：
                   −2147483647 取反得 +2147483647，可表且正确，属正常路径；
                   真正不可表的只有 −2147483648 这一个值，故只有它落饱和出口；
                ④ 饱和时返回正向毫秒上限并升故障级——调用方必须知道这个幅值是钳位值；
                ⑤ 负输入取到幅值后发信息级并置 bNegative，方向信息不丢。
                职责边界：带偏移的时刻算术归 FC_DL_TodAddWrap / FC_DL_TodDiffWrap；
                TIME 与秒的换算归 FC_DL_TimeToLrealSec / FC_DL_LrealSecToTime；
                本件只管「幅值」这一件事。
    编译门槛  : 主路径假设 TIME 以 32 位毫秒（DINT）承载，CODESYS V3.5+ / TwinCAT 3 /
                InoProShop 均为该口径。若目标平台 TIME 为 64 位容器，TIME_TO_DINT 会在
                超出 32 位时截断——此时应改用 64 位换算链，本件的闸门顺序与出口不变。
                饱和值以 DINT 常量经 DINT_TO_TIME 落地，不使用超长 TIME 字面量，
                避免 32 位 TIME 平台上字面量本身无法编译。
    错误码    : 16#0001_042E 输入为负，已取绝对值（bNegative 可查）——信息级，值可用
                16#0001_042F 预留禁用（信息级，不得挪用）
                16#0001_0363 −MAX−1 的绝对值不可用 DINT 表达，已饱和至正向上限——故障级，bValid = FALSE
                16#0001_0364 预留（故障级，不得挪用）
                16#0001_0365 预留禁用（故障级，不得挪用）
    码位总账  : 16#0001_042E 用 / 16#0001_042F 预留 ｜ 16#0001_0363 用 / 16#0001_0364 预留 / 16#0001_0365 预留
    状态机    : R6 标注 N/A —— 本组件为纯函数无顺序状态机，无 CASE 可写，非法状态不可能出现
    采样约定  : 本件无定时器、无沿检测、无状态；单拍纯计算，结论与任务周期无关。
    修订记录  : 2026-11-16 v1.0.0 首次入库（R20）
*)
FUNCTION FC_DL_TimeAbsSat : TIME
VAR_INPUT
    tIn              : TIME;                  // 输入时长，可负 [ms]，TIME 平台实现为 32 位毫秒 / input duration, signed [ms], TIME is 32-bit milliseconds on the target platforms
END_VAR
VAR_OUTPUT
    eErr             : UDINT;                 // 错误码，0=正常 / error id, 0=ok
    bError           : BOOL;                  // 故障标志，eErr 为故障级时 TRUE / error flag, TRUE on fault-level eErr
    bValid           : BOOL;                  // 返回值是否可用（饱和时为 FALSE）/ return usable, FALSE when saturated
    bNegative        : BOOL;                  // 输入为负，已取绝对值 / the input was negative and its magnitude is published
END_VAR
VAR CONSTANT
    DL_TIME_MS_POS_MAX : DINT := 2147483647;  // DINT 毫秒正向上限，饱和出口值 [ms] / DINT millisecond top, the saturation value [ms]
    DL_TIME_MS_NEG_SAFE : DINT := -2147483647; // 可安全取负的毫秒下界，即 −MAX [ms] / the lowest value that can be negated safely, minus MAX [ms]
    DL_DINT_ZERO     : DINT := 0;             // 有符号零常量，避免裸字面量 [ms] / signed zero constant [ms]
    DL_TIME_ZERO     : TIME := T#0s;          // 零时长，缺省返回 / zero duration returned by default
END_VAR
VAR
    nIn              : DINT;                  // 输入毫秒中间量 [ms] / input milliseconds intermediate [ms]
    nAbs             : DINT;                  // 绝对值毫秒中间量 [ms] / magnitude intermediate in milliseconds [ms]
END_VAR

// 段 1｜返回值与错误状态预置 / segment 1, preset return value and error status
FC_DL_TimeAbsSat := DL_TIME_ZERO;             // 缺省返回零时长 / default returns a zero duration
eErr := 0;                                    // 预置无错误 / preset no error
bError := FALSE;                              // 预置无故障 / preset no fault
bValid := FALSE;                              // 预置不可用，通过闸门后置位 / preset invalid, set TRUE after the gates
bNegative := FALSE;                           // 预置输入非负 / preset a non-negative input
nAbs := DL_DINT_ZERO;                         // 幅值中间量清零 / clear the magnitude intermediate

// 段 2｜取值：显式标准转换，禁隐式 / segment 2, explicit standard conversion, never implicit
nIn := TIME_TO_DINT(tIn);                     // TIME → 毫秒 [ms] / TIME to milliseconds [ms]

// 段 3｜非负直通：幅值即原值，零开销 / segment 3, non-negative pass-through with zero overhead
IF nIn >= DL_DINT_ZERO THEN
    FC_DL_TimeAbsSat := DINT_TO_TIME(nIn);    // 幅值即原值 [ms] / the magnitude is the value itself [ms]
    bValid := TRUE;                           // 直通值可用 / the pass-through value is usable
    RETURN;                                   // 出口 / exit
END_IF

// 段 4｜−MAX−1 边界闸：相反数不可表，先判后算 / segment 4, the unrepresentable boundary gate
IF nIn < DL_TIME_MS_NEG_SAFE THEN
    FC_DL_TimeAbsSat := DINT_TO_TIME(DL_TIME_MS_POS_MAX); // 饱和至正向毫秒上限 [ms] / saturate to the positive millisecond top [ms]
    eErr := 16#0001_0363;                     // 故障级：−MAX−1 的绝对值不可表达 / fault level, the magnitude of minus MAX minus one is not representable
    bError := TRUE;                           // 置故障标志 / raise the error flag
    bValid := FALSE;                          // 饱和值不可作统计依据 / the saturated value must not feed the statistics
    bNegative := TRUE;                        // 输入确实为负 / the input really was negative
    RETURN;                                   // 出口 / exit
END_IF

// 段 5｜正常负值取幅值（此处取反结构性安全：nIn 严格大于可安全下界）/ segment 5, negate a safe negative value
nAbs := -nIn;                                 // 取绝对值 [ms] / take the magnitude [ms]
FC_DL_TimeAbsSat := DINT_TO_TIME(nAbs);       // 回装为时长 [ms] / convert back into a duration [ms]
eErr := 16#0001_042E;                         // 信息级：输入为负，已取绝对值 / info level, the negative input was turned into a magnitude
bNegative := TRUE;                            // 方向信息不丢 / the direction information is kept
bValid := TRUE;                               // 幅值可用 / the magnitude is usable
END_FUNCTION

(* ---- FC_DL_TimeAddSat.st ---- *)
(*
    FC_DL_TimeAddSat —— TIME 加法溢出饱和防御包装
    ------------------------------------------------------------------
    分类      : DL_MathData / TimeArith
    前缀      : FC_DL_
    版本      : 1.0.0
    溯源      : IEC 61131-3 标准语义的道莅防御性实现
                （内部委托平台内建函数，外围统一错误码/钳位/双语文档；
                  未复制任何闭源厂商源码，参考实现仅限 MIT/Apache 许可）
    平台      : 纯 IEC 61131-3，CODESYS / TwinCAT / InoProShop 通用
    作者      : 道莅代码库 · PLC编程专家（R16）
    ------------------------------------------------------------------
    功能说明  : TIME 加法：返回 tA + tB，TIME 算术委托 `+` 与 `-` 运算符，
                不重实现任何时间运算内核；
                溢出预判采用减法比较口径（规避「先算后判」红线）：
                tA > DL_TIME_MAX - tB 时判加法将溢出，直接饱和输出 DL_TIME_MAX，
                置信息级 16#0001_01E0（bError=FALSE、bValid=TRUE）；
                预判安全性：TIME 为 32 位无符号容器，tB 恒 ≤ DL_TIME_MAX，
                故 DL_TIME_MAX - tB 恒 ≥ T#0S，减法比较本身不下溢；
                钳位方向：仅上界单侧饱和至 DL_TIME_MAX（T#49D17H2M47S295MS）；
                常量字面量说明：DL_TIME_MAX 采用 D/H/M/S/MS 组合字面量（三大平台均支持），
                等价于 ms 口径 4294967295 ms，若目标平台不支持组合字面量可改为 T#4294967295MS。
    错误码    : 16#0001_01E0 加法结果超 TIME 上限，已饱和至 DL_TIME_MAX——信息级，正常防御
                16#0001_01E1 预留禁用（信息级，不得挪用）
                16#0001_02BE 预留禁用（故障级，不得挪用）
                16#0001_02BF 预留禁用（故障级，不得挪用）
                16#0001_02C0 预留禁用（故障级，不得挪用）
    状态机    : R6 标注 N/A —— 本组件为纯函数无顺序状态机，无 CASE 可写，非法状态不可能出现，故以本节说明替代 ELSE 兜底
    修订记录  : 2026-11-16 v1.0.0 首次入库（R16）
*)
FUNCTION FC_DL_TimeAddSat : TIME
VAR_INPUT
    tA : TIME; // 加数 A [ms] / addend A
    tB : TIME; // 加数 B [ms] / addend B
END_VAR
VAR_OUTPUT
    eErr   : UDINT; // 错误码，0=正常 / error id, 0=ok
    bError : BOOL;  // 是否出错，eErr 非 0 时为 TRUE / error flag, TRUE when eErr is nonzero
    bValid : BOOL;  // 输出是否有效可用 / output valid flag
END_VAR
VAR CONSTANT
    DL_TIME_MAX   : TIME := T#49D17H2M47S295MS; // 32 位 TIME 容器上限，等价 4294967295 ms [ms] / 32-bit TIME container ceiling, equals 4294967295 ms
    DL_TIME_ZERO  : TIME := T#0S;               // TIME 零值 [ms] / TIME zero value
END_VAR

// 段 1｜返回值与错误状态预置 / segment 1, preset return value and error status
FC_DL_TimeAddSat := DL_TIME_ZERO; // 故障缺省返回 T#0S [ms] / fault default returns T#0S
eErr   := 0;     // 预置无错误 / preset no error
bError := FALSE; // 预置无故障 / preset no fault
bValid := FALSE; // 预置无效，通过溢出预判后置位 / preset invalid, set TRUE after overflow pre-check

// 段 2｜减法比较溢出预判与主体加法（末段） / segment 2, subtract-compare overflow pre-check and main addition (final)
IF tA > DL_TIME_MAX - tB THEN
    FC_DL_TimeAddSat := DL_TIME_MAX; // 溢出预判命中，饱和至上限（tB ≤ DL_TIME_MAX 恒成立，预判减法不下溢） / overflow pre-check hit, saturate to ceiling (tB never exceeds DL_TIME_MAX, pre-check subtraction cannot underflow)
    eErr := 16#0001_01E0;            // 信息级：加法溢出已饱和 / info level: addition overflow, saturated
ELSE
    FC_DL_TimeAddSat := tA + tB; // 预判通过，域内委托 `+` 运算符加法 / pre-check passed, in-domain addition via `+` operator
    eErr := 0; // 域内无错误 / in-domain, no error
END_IF
bError := FALSE; // 信息级饱和不置故障 / info-level saturation never raises fault
bValid := TRUE;  // 域内或饱和输出均有效可用 / in-domain or saturated output is valid
END_FUNCTION

(* ---- FC_DL_TimeClampEx.st ---- *)
(*
    FC_DL_TimeClampEx —— TIME 三参钳制（跨平台 LIMIT 等价实现）
    ------------------------------------------------------------------
    分类      : DL_MathData / TimeArith
    前缀      : FC_DL_
    版本      : 1.0.0
    溯源      : IEC 61131-3 标准语义的道莅防御性实现
                （LIMIT(MN, IN, MX) 的 TIME 版本；部分平台只对数值类型定义
                  LIMIT / MAX / MIN，对 TIME 未定义或不接受混型实参，故以纯比较式
                  等价实现，禁用任何平台内建 LIMIT，保证四平台行为逐字一致；
                  clean-room 编写，未复制任何闭源厂商源码）
    平台      : 纯 IEC 61131-3，CODESYS 3.5 / TwinCAT 3 / InoProShop / Machine Expert 通用
    作者      : 道莅代码库 · PLC编程专家（R69 构建轮 · 批 1 · N2）
    ------------------------------------------------------------------
    功能说明  : 把时长钳在 [tMin, tMax] 闭区间内。跨平台口径说明（这是本件存在的
                唯一理由）：IEC 61131-3 对 LIMIT 只给出数值类型形式，TIME 实参在
                CODESYS 上可编译而在部分平台直接报「不支持的类型组合」，现场
                换平台时同一行代码从「可编译」变成「编译失败」，属不可移植风险。
                本件以两条比较改写，语义与 LIMIT 逐字等价：
                IN < MN -> MN ；IN > MX -> MX ；区间内直通。
                区间序闸：tMin > tMax 视为组态非法（区间退化 / 反向），**禁入**并
                报故障级；故障缺省返回 tMin（安全侧：钳制件的安全端是下限，避免
                把「区间填反」放大成「超长保持」）。tMin = tMax 是合法退化区间
                （退化为定值），不报码。
                越界钳位报信息级（值可用），区间内直通不报码。
    错误码    : 16#0001_03F9 钳位区间非法（tMin > tMax），输出 tMin —— 故障级
                16#0001_04F7 输入越界已被钳制（bClamped 可查）—— 信息级，值可用
    码位总账  : 16#0001_03F9 用 ｜ 16#0001_04F7 用
    状态机    : R6 标注 N/A —— 纯函数无顺序状态机，无 CASE 可写，非法状态不可能出现
    采样约定  : 无定时器 / 无沿检测 / 无跨周期状态，结论与任务周期无关
    修订记录  : 2026-11-22 v1.0.0 首次入库（R69 构建轮 · 批 1 · N2）
*)
FUNCTION FC_DL_TimeClampEx : TIME
VAR_INPUT
    tIn   : TIME;                              // 待钳制时长 [ms] / duration to clamp [ms]
    tMin  : TIME;                              // 区间下限（含） [ms] / lower bound, inclusive [ms]
    tMax  : TIME;                              // 区间上限（含） [ms] / upper bound, inclusive [ms]
END_VAR
VAR_OUTPUT
    eErr     : UDINT;                          // 错误码，0 = 正常 / error id, 0 = ok
    bError   : BOOL;                           // 故障标志，仅故障级码置 TRUE / error flag, TRUE on fault level only
    bValid   : BOOL;                           // 返回值可用（故障级为 FALSE）/ return usable, FALSE on fault level
    bClamped : BOOL;                           // 本次发生了钳制 / a clamp actually happened
END_VAR
VAR CONSTANT
    DL_TC_ZERO : TIME := T#0S;                 // TIME 零值常量（占位，不参与钳制） [ms] / TIME zero constant
END_VAR

// 段 1｜返回值与错误状态预置（实战规则 1①）/ segment 1, preset the return value and the status
FC_DL_TimeClampEx := DL_TC_ZERO;   // 缺省返回 T#0S，过闸后按分支覆盖 [ms] / default T#0S, overwritten below
eErr     := 0;                     // 预置无错误 / preset no error
bError   := FALSE;                 // 预置无故障 / preset no fault
bValid   := FALSE;                 // 预置不可用 / preset unusable
bClamped := FALSE;                 // 预置未钳制 / preset unclamped

// 段 2｜区间序闸：tMin > tMax 属组态非法，禁入（安全侧返回下限）/ segment 2, interval order gate
IF tMin > tMax THEN
    FC_DL_TimeClampEx := tMin;     // 安全侧返回下限，绝不把反向区间放大成超长值 [ms] / safe side returns the lower bound
    eErr   := 16#0001_03F9;        // 故障级：钳位区间非法 / fault level: illegal clamp interval
    bError := TRUE;                // R45 配对 / paired with the code
    bValid := FALSE;               // 返回值不可用 / return unusable
    RETURN;                        // 出口 / exit
END_IF

// 段 3｜钳制主体：两条比较改写，语义与 LIMIT(MN, IN, MX) 逐字等价 / segment 3, clamp body
IF tIn < tMin THEN
    FC_DL_TimeClampEx := tMin;     // 低于下限：钳到下限 [ms] / below the floor, clamp up
    bClamped := TRUE;              // 钳制发生 / clamp happened
    eErr     := 16#0001_04F7;      // 信息级：输入越界已钳制 / info level: input out of range, clamped
ELSIF tIn > tMax THEN
    FC_DL_TimeClampEx := tMax;     // 高于上限：钳到上限 [ms] / above the ceiling, clamp down
    bClamped := TRUE;              // 钳制发生 / clamp happened
    eErr     := 16#0001_04F7;      // 信息级：输入越界已钳制 / info level: input out of range, clamped
ELSE
    FC_DL_TimeClampEx := tIn;      // 区间内（含两端）直通 [ms] / inside the interval, pass through
END_IF

bError := FALSE;   // 信息级钳制不置故障（钳制是防御而非故障）/ info-level clamping is a defence, not a fault
bValid := TRUE;    // 三条分支的输出均可用 / usable in all three branches
END_FUNCTION
